(* IEC 61131-3 sources: daoli-st-library/DL_Process (part 50) *)

(* ---- FB_DL_SampleLoopPurge.st ---- *)
(*
  FB_DL_SampleLoopPurge  —  取样回路吹扫与取样窗（阀序 + 吹扫/静置计时） / Sample-loop purge and sampling window with valve sequence and purge/settle timers
  分类 Category : DL_Process
  版本 Version  : 1.0.0
  来源 Source   : t1-2-oscat-building — 楼宇/工艺分析取样回路阀序族深化
  溯源 Origin   : 道莅 clean-room 实现；吹扫-静置-取样三段阀序与计时为公开取样系统工艺逻辑，未复制任何源码行
  功能 Function : 1) 三段阀序：ePurge 吹扫（吹扫阀开 + 需 bFlowOk 有流，tPurge 到时）→
                  eSettle 静置（全阀关，tSettle 到时）→ eSample 取样窗（取样阀开，tSample 到时）→
                  eDone；2) 吹扫超时（无流）判故障；3) 取样窗内 bSampleReady 丢失判故障；
                  4) 故障级单码 03A4，归因由 eCause 独立成员承载（R190）；
                  5) 信息级 04CC = 取样窗完成沿；6) 解除式全当拍量（R240）。
  接口 Interface: 输入有流/取样就绪/三个时间量；输出状态 + 三阀位 + 码
  边界 Boundary : ① 组态闸：三个时间量 <= T#0S 任一成立 → 03A4 锁存；
                  ② 三阀位由相位单点映射（段 6），故障相全阀关断（安全侧）；
                  ③ 三个 TON 段 0 无条件周期调用，IN 由相位派生，相切换自动复位 ET（R176）；
                  ④ 取样窗内就绪丢失为「事件消失」判据，非单拍标志门控（禁 bError 门控）；
                  ⑤ 故障相迁出唯一路径 = bReset 上升沿；⑥ 零全局耦合（无 GVL / %I %Q %M）。
  依赖 Depends  : Standard.library（TON / R_TRIG）
  码表 Error codes（Process 段 0005，故障窗口 03A4 / 信息窗口 04CC）:
    16#0005_03A4 故障级：取样回路故障总码（组态非法 / 吹扫超时无流 / 取样窗就绪丢失），
                 锁存至 bReset 上升沿；归因见 eCause，不新增码位（派单硬约束单码）
    16#0005_04CC 信息级：取样窗完成沿（进 eDone 单拍）
  修订历史 Revision :
    2026-11-19  v1.0.0  R43 首版（批次 2 · 序号 8）
*)

TYPE E_DL_SlpState :
(
    eIdle   := 0,     // 未使能：全阀关 / Idle, all valves closed
    ePurge  := 10,    // 吹扫中 / Purging
    eSettle := 20,    // 静置中（全阀关） / Settling with valves closed
    eSample := 30,    // 取样窗中 / Sampling window
    eDone   := 50,    // 循环完成 / Done
    eFault  := 90     // 故障锁存相（全阀关） / Fault latched, valves closed
);
END_TYPE

TYPE E_DL_SlpCause :
(
    eNone       := 0, // 无故障成因 / No cause
    eCfgIllegal := 1, // 组态非法 / Illegal configuration
    ePurgeTmo   := 2, // 吹扫超时无流 / Purge timeout without flow
    eSampleLost := 3  // 取样窗就绪丢失 / Sampling readiness lost
);
END_TYPE

FUNCTION_BLOCK FB_DL_SampleLoopPurge
VAR_INPUT
    bFlowOk      : BOOL := FALSE;      // 吹扫有流反馈（电平）[-] / Purge flow feedback
    bSampleReady : BOOL := FALSE;      // 取样就绪（电平）[-] / Sampling ready
    tPurge       : TIME := T#30S;      // 吹扫时长 [ms]，域 > 0 / Purge duration
    tSettle      : TIME := T#5S;       // 静置时长 [ms]，域 > 0 / Settle duration
    tSample      : TIME := T#10S;      // 取样窗时长 [ms]，域 > 0 / Sampling window
    bStart       : BOOL := FALSE;      // 启动命令（电平）[-] / Start command
    bReset       : BOOL := FALSE;      // 复位命令，上升沿清故障 [-] / Reset edge
END_VAR
VAR_OUTPUT
    eState       : E_DL_SlpState;      // 状态出口，段 6 单点映射 / State outlet
    eCause       : E_DL_SlpCause;      // 故障成因出口（R190） / Fault cause outlet
    bPurgeValve  : BOOL;               // 吹扫阀指令 [-] / Purge valve command
    bSampleValve : BOOL;               // 取样阀指令 [-] / Sample valve command
    bVentValve   : BOOL;               // 排放阀指令 [-] / Vent valve command
    bCycleDone   : BOOL;               // 循环完成标志 [-] / Cycle done flag
    bError       : BOOL;               // 故障锁存标志 [-] / Fault latch flag
    nErrId       : UDINT;              // 事件码，0 = 无事件 / Event code
END_VAR
VAR
    _eState      : E_DL_SlpState := E_DL_SlpState.eIdle;   // 内部相位（CASE 唯一写入目标） / Internal phase
    _eCause      : E_DL_SlpCause := E_DL_SlpCause.eNone;   // 故障成因锁存（锁存量） / Latched cause
    tonPurge     : TON;                // 吹扫计时，每周期无条件调用 / Purge timer
    tonSettle    : TON;                // 静置计时，每周期无条件调用 / Settle timer
    tonSample    : TON;                // 取样窗计时，每周期无条件调用 / Sampling timer
    rtReset      : R_TRIG;             // 复位沿实例，每周期无条件调用 / Reset edge
    _bCfgBad     : BOOL;               // 组态非法当拍量 [-] / Config illegal
    _bFault      : BOOL;               // 故障锁存位（锁存量） / Latched fault bit
    _uFault      : UDINT;              // 故障码锁存（锁存量） / Latched fault code
    _uInfo       : UDINT;              // 信息码，每拍重算 / Transient info code
END_VAR

(* —— 段 0：沿实例与定时器无条件周期刷新（IN 由相位派生，相内自动清零 ET） —— *)
_bCfgBad := (tPurge <= T#0S) OR (tSettle <= T#0S) OR (tSample <= T#0S);     // 组态非法当拍量 / Config illegal
rtReset(CLK := bReset);                                                     // 复位沿，每拍必调 / Reset edge
tonPurge(IN := (_eState = E_DL_SlpState.ePurge), PT := tPurge);             // 吹扫计时 / Purge timer
tonSettle(IN := (_eState = E_DL_SlpState.eSettle), PT := tSettle);          // 静置计时 / Settle timer
tonSample(IN := (_eState = E_DL_SlpState.eSample), PT := tSample);          // 取样窗计时 / Sampling timer

(* —— 段 1：单拍量预清零（锁存量不入清单） —— *)
_uInfo := 16#0000_0000;            // 信息码每拍重算 / Info recomputed
bPurgeValve := FALSE;              // 吹扫阀缺省关 / Purge valve default closed
bSampleValve := FALSE;             // 取样阀缺省关 / Sample valve default closed
bVentValve := FALSE;               // 排放阀缺省关 / Vent valve default closed
bCycleDone := FALSE;               // 完成标志缺省 FALSE / Done default
nErrId := 16#0000_0000;            // 事件码缺省无事件 / Event code default

(* —— 段 2：复位沿 + 组态域闸 —— *)
IF rtReset.Q THEN                              // rtReset.Q = 当拍量 / current scan
    _bFault := FALSE;                          // 清故障锁存位（锁存量） / Clear fault latch
    _uFault := 16#0000_0000;                   // 清故障锁存码（锁存量） / Clear fault code
    _eCause := E_DL_SlpCause.eNone;            // 清成因（锁存量） / Clear cause
    IF _eState = E_DL_SlpState.eFault THEN
        _eState := E_DL_SlpState.eIdle;        // 故障相迁出：回未使能 / Fault exit to idle
    END_IF
END_IF
IF _bCfgBad THEN                               // 组态域闸 / Config gate
    _uFault := 16#0005_03A4;                   // 故障级：取样回路故障总码 / Process fault code
    _eCause := E_DL_SlpCause.eCfgIllegal;      // 归因：组态非法 / Cause: illegal config
    _bFault := TRUE;                           // 标志与码位配对（R45） / Flag paired with code
END_IF

(* —— 段 3：吹扫超时无流 / 取样窗就绪丢失（判据当拍量） —— *)
IF (NOT _bFault) AND (_eState = E_DL_SlpState.ePurge) AND (NOT bFlowOk) THEN
    _uFault := 16#0005_03A4;
    _eCause := E_DL_SlpCause.ePurgeTmo;        // 归因：吹扫无流 / Cause: purge without flow
    _bFault := TRUE;
END_IF
IF (NOT _bFault) AND (_eState = E_DL_SlpState.eSample) AND (NOT bSampleReady) THEN
    _uFault := 16#0005_03A4;
    _eCause := E_DL_SlpCause.eSampleLost;      // 归因：取样就绪丢失 / Cause: readiness lost
    _bFault := TRUE;
END_IF

(* —— 段 4：故障解除式（R240；全当拍量）：rtReset.Q / NOT _bCfgBad / NOT tonPurge.Q / bFlowOk —— *)
IF rtReset.Q AND (NOT _bCfgBad) AND (NOT tonPurge.Q) THEN
    _bFault := FALSE;                          // 清故障锁存位（锁存量） / Clear fault latch
    _uFault := 16#0000_0000;                   // 清故障锁存码（锁存量） / Clear fault code
    _eCause := E_DL_SlpCause.eNone;            // 清成因（锁存量） / Clear cause
END_IF

(* —— 段 4A：故障锁存相位迁移闸 —— *)
IF _bFault AND (_eState <> E_DL_SlpState.eFault) THEN
    _eState := E_DL_SlpState.eFault;           // 锁存即入故障相（全阀关） / Latch enters fault phase
END_IF

(* —— 段 5：相位机（CASE 全覆盖 + ELSE 兜底） —— *)
CASE _eState OF

E_DL_SlpState.eIdle:
    IF bStart AND (NOT _bFault) THEN           // 启动条件 / Start gate
        _eState := E_DL_SlpState.ePurge;       // 进吹扫相 / Enter purge
    END_IF

E_DL_SlpState.ePurge:
    bPurgeValve := TRUE;                       // 吹扫阀开 / Purge valve open
    bVentValve := TRUE;                        // 排放阀开（吹扫排空） / Vent valve open
    IF tonPurge.Q AND bFlowOk THEN             // 出口 1：吹扫到时且有流 / Purge done with flow
        _eState := E_DL_SlpState.eSettle;      // 进静置相 / Enter settle
    ELSIF NOT bStart THEN                      // 出口 2：撤启动（R98 双出口） / Start released
        _eState := E_DL_SlpState.eIdle;
    END_IF

E_DL_SlpState.eSettle:
    IF tonSettle.Q THEN                        // 静置到时（全阀关） / Settle elapsed
        _eState := E_DL_SlpState.eSample;      // 进取样窗 / Enter sampling
    ELSIF NOT bStart THEN                      // 撤启动：中止 / Abort
        _eState := E_DL_SlpState.eIdle;
    END_IF

E_DL_SlpState.eSample:
    bSampleValve := TRUE;                      // 取样阀开 / Sample valve open
    IF tonSample.Q THEN                        // 取样窗到时 / Sampling elapsed
        _uInfo := 16#0005_04CC;                // 信息级：取样窗完成沿 / Info: sampling complete
        _eState := E_DL_SlpState.eDone;        // 进完成相 / Enter done
    ELSIF NOT bStart THEN                      // 撤启动：中止 / Abort
        _eState := E_DL_SlpState.eIdle;
    END_IF

E_DL_SlpState.eDone:
    IF NOT bStart THEN                         // 撤启动回空闲 / Start released returns idle
        _eState := E_DL_SlpState.eIdle;
    END_IF

E_DL_SlpState.eFault:
    ;                                          // 故障相：全阀关断，仅段 4 复位沿可迁出 / Valves closed, reset only

ELSE
    _uFault := 16#0005_03A4;                   // 故障级：非法相位兜底（归并总码） / Illegal phase fallback
    _eCause := E_DL_SlpCause.eCfgIllegal;      // 归因：相位非法归并组态 / Cause: phase illegal
    _bFault := TRUE;
    _eState := E_DL_SlpState.eFault;           // 强制回故障相 / Force fault phase

END_CASE

(* —— 段 6：出口单点映射（名实同源；故障相全阀关断为安全侧） —— *)
IF _bFault THEN
    bPurgeValve := FALSE;                      // 故障相吹扫阀强制关 / Purge valve forced closed
    bSampleValve := FALSE;                     // 故障相取样阀强制关 / Sample valve forced closed
    bVentValve := FALSE;                       // 故障相排放阀强制关 / Vent valve forced closed
    nErrId := _uFault;                         // 故障锁存码回放 / Replay latched code
ELSE
    nErrId := _uInfo;                          // 信息码 / Transient info
END_IF
bCycleDone := (_eState = E_DL_SlpState.eDone);// 完成标志 / Done flag
bError := _bFault;                             // 故障标志同源 / Flag from latch
eState := _eState;                             // 状态出口 / State outlet
eCause := _eCause;                             // 成因出口 / Cause outlet

END_FUNCTION_BLOCK

(* ---- FB_DL_ScreenPanelWearMonitor.st ---- *)
(*
  Name: FB_DL_ScreenPanelWearMonitor
  Category: DL_Process
  Version: 1.0.0
  Round: R89 / 2026-11-25
  开源溯源：clean-room 自研（族 矿山破碎筛分，ST 开源生态实测 0 命中，无外部代码引入）
  功能：筛板磨损监测（累计过料量法）：按运行时间积分过料吨位，乘磨损系数得累计磨损厚度与剩余寿命。
  边界条件：① 五浮点入参全部过非有限闸，任一非有限进冻结分支：输出保持上一有效值 + xValid = FALSE；
            ② 累计量为跨拍保持量，首扫以 _bInit 初始化，xReset 只清累计吨位（作用域：清累计，不清配置）；
            ③ 周期换算口径：TIME_TO_REAL 取毫秒（库内统一口径），tCycleS ≤ 0 时以 10 ms 缺省兜底；
            ④ 磨损厚度饱和于有效厚度差（钳的是剩余寿命量值，xValid 不受影响）。
  量纲自证：fFeedTph[t/h] × dt[h] = t；t/1000 = kt；kt × fWearCoef[mm/kt] = mm。
*)
FUNCTION_BLOCK FB_DL_ScreenPanelWearMonitor
VAR_INPUT
    xRun : BOOL;                (* 筛机运行反馈 [-] Screen running *)
    fFeedTph : REAL;            (* 瞬时给料量 [t/h] Instantaneous feed rate [t/h] *)
    fWearCoef : REAL;           (* 磨损系数 [mm/kt] Wear coefficient [mm per kilotonne] *)
    fPanelThkInitMm : REAL;     (* 筛板初始厚度 [mm] Initial panel thickness [mm] *)
    fPanelThkMinMm : REAL;      (* 筛板报废厚度 [mm] Scrap thickness [mm] *)
    xReset : BOOL;              (* 累计清零（换板后置位一拍） [-] Reset accumulation *)
    tCycleS : TIME;             (* 扫描周期 [ms] Scan cycle [ms] *)
END_VAR
VAR_OUTPUT
    fWornMm : REAL;             (* 累计磨损厚度 [mm] Accumulated wear [mm] *)
    fRemainLifePct : REAL;      (* 剩余寿命百分比 [%] Remaining life [%] *)
    xReplaceAlarm : BOOL;       (* 换板报警（剩余 ≤ 10 %） [-] Replace alarm *)
    xValid : BOOL;              (* 配置与链路有效 [-] Configuration and chain valid *)
END_VAR
VAR
    _bInit : BOOL := FALSE;     (* 首扫初始化标志 [-] First-scan init flag *)
    _bCfgBad : BOOL := FALSE;   (* 配置非法当拍量 [-] Configuration bad *)
    _bCalcOk : BOOL := FALSE;   (* 本拍计算有效 [-] Calculation valid this scan *)
    _fTonsAcc : REAL := 0.0;    (* 累计过料量 [t] Accumulated tonnage [t] *)
    _fWorn : REAL := 0.0;       (* 累计磨损厚度保持量 [mm] Wear thickness hold [mm] *)
    _fRemain : REAL := 0.0;     (* 剩余寿命保持量 [%] Remaining life hold [%] *)
    _fSpanMm : REAL := 0.0;     (* 有效可磨损厚度差 [mm] Usable thickness span [mm] *)
    _fDtH : REAL := 0.0;        (* 本拍时间步长 [h] Time step [h] *)
END_VAR
VAR CONSTANT
    DL_EPS : REAL := 1.0E-9;        (* 除零判定容差 [-] Divide-by-zero tolerance *)
    DL_KT : REAL := 1000.0;         (* 吨 → 千吨换算 [t/kt] Tonne to kilotonne *)
    DL_SECH : REAL := 3600.0;       (* 秒 → 小时换算 [s/h] Second to hour *)
    DL_CYCDEF : REAL := 0.01;       (* 缺省扫描周期 [s] Default scan cycle [s] *)
    DL_ALARM_PCT : REAL := 10.0;    (* 换板报警门限（剩余寿命） [%] Replace alarm threshold [%] *)
    DL_PCT : REAL := 100.0;         (* 百分数基准 [%] Percent base *)
END_VAR
(* 首扫初始化：累计量与保持量一次性归零（R310） *)
IF NOT _bInit THEN
    _fTonsAcc := 0.0;
    _fWorn := 0.0;
    _fRemain := DL_PCT;
    _bInit := TRUE;
END_IF
(* 周期换算：毫秒 → 秒 → 小时；非正周期以缺省 10 ms 兜底 *)
IF tCycleS <= T#0S THEN
    _fDtH := DL_CYCDEF / DL_SECH;
ELSE
    _fDtH := (TIME_TO_REAL(tCycleS) / 1000.0) / DL_SECH;
END_IF
(* 复位作用域：只清累计吨位与磨损量，不动配置与报警门限 *)
IF xReset THEN
    _fTonsAcc := 0.0;
    _fWorn := 0.0;
    _fRemain := DL_PCT;
END_IF
(* 非有限闸（NaN 自反 + Inf 差值自减）+ 组态域闸：五浮点入参全枚举（R272） *)
_bCfgBad := (fFeedTph <> fFeedTph) OR ((fFeedTph - fFeedTph) <> 0.0)
         OR (fWearCoef <> fWearCoef) OR ((fWearCoef - fWearCoef) <> 0.0)
         OR (fPanelThkInitMm <> fPanelThkInitMm) OR ((fPanelThkInitMm - fPanelThkInitMm) <> 0.0)
         OR (fPanelThkMinMm <> fPanelThkMinMm) OR ((fPanelThkMinMm - fPanelThkMinMm) <> 0.0)
         OR (fFeedTph < 0.0) OR (fFeedTph > 5000.0)
         OR (fWearCoef < 0.0) OR (fWearCoef > 20.0)
         OR (fPanelThkMinMm <= 0.0) OR (fPanelThkInitMm <= (fPanelThkMinMm + DL_EPS))
         OR (fPanelThkInitMm > 200.0);
_bCalcOk := NOT _bCfgBad;
IF _bCalcOk THEN
    (* 运行中按周期积分过料吨位：t/h × h = t *)
    IF xRun THEN
        _fTonsAcc := _fTonsAcc + fFeedTph * _fDtH;
    END_IF
    (* 累计磨损厚度：t → kt，kt × [mm/kt] = mm *)
    _fWorn := (_fTonsAcc / DL_KT) * fWearCoef;
    (* 剩余寿命：有效厚度差已过正性闸，绝无零除 *)
    _fSpanMm := fPanelThkInitMm - fPanelThkMinMm;
    _fRemain := (1.0 - _fWorn / _fSpanMm) * DL_PCT;
    (* 极限钳位：磨穿即 0 %，新板不超 100 % *)
    IF _fWorn >= _fSpanMm THEN
        _fRemain := 0.0;
    END_IF
    IF _fRemain < 0.0 THEN
        _fRemain := 0.0;
    ELSIF _fRemain > DL_PCT THEN
        _fRemain := DL_PCT;
    END_IF
END_IF
(* 统一出口（单点赋值）：冻结分支保持上一有效值，保持量来源均为已过闸的有限值（R273） *)
fWornMm := _fWorn;
fRemainLifePct := _fRemain;
xReplaceAlarm := _bCalcOk AND (_fRemain <= DL_ALARM_PCT);
xValid := _bCalcOk;
END_FUNCTION_BLOCK

(* ---- FB_DL_ScrewPressDewaterSeq.st ---- *)
(*
  道莅工业代码库 / Daoli Industrial ST Library
  组件: FB_DL_ScrewPressDewaterSeq
  分类: DL_Process
  复杂度: C4 ｜ 版本: 1.0.0 ｜ 2026-11-24
  平台兼容: CODESYS 3.5+ / TwinCAT 3 / 汇川 InoProShop / 施耐德 Machine Expert
  开源溯源: 无（clean-room 工程时序自研；参考公开的螺旋压榨脱水机单循环工艺步骤，
            未复制任何受版权保护代码）
  许可证: 本项目自有 (MIT)

  功能职责:
    污泥螺旋压榨脱水机单循环时序：进泥 → 加药混合 → 压榨 → 冲洗 → 退让复位。
    互锁：eFeed 要求 bFeedOk AND bPolyOk（缺料进故障码 21）；ePress 期间 bPressHigh
    累计超过 tPress 的 30% 即提前转 eFlush（过压保护，码 22，先降后报的安全侧）；
    bPressFault 任意相进故障码 23 并在同一拍切断 bPressMotor；bStop 任意相转 eRetract（码 26）。

  输入/输出契约:
    IN  bStart 上升沿启动；bStop 任意相转退让相；bReset 上升沿是 eFault 唯一出口。
    OUT 四个执行输出全部为「单稳态、每拍按相位重算、不锁存」，eFault 内全部 FALSE。

  码表 (Codes):
    21 = 进泥或加药未就绪（故障级；转 eFault）
    22 = 压榨过压提前转冲洗（降级级安全侧；不置故障相）
    23 = 压榨机故障（故障级；同拍断 bPressMotor）
    24 = 泥饼含固率低于设定（信息级；本循环照常结束，仅记录）
    25 = 泥饼含固率信号非有限（故障级）
    26 = 停止指令触发退让（信息级）
    27 = 时间参数越域且不满足 tPress > tMix（故障级；约束不成立则过压窗口无意义）
    28 = 过压触发次数达上限（故障级；同一循环内反复过压视为机械异常）
    99 = 非法状态枚举值（ELSE 兜底）

  边界与红线:
    ① 六个 TON 与两个 R_TRIG 全在 CASE 外无条件刷新（R7），CASE 内只读 .Q / .ET。
    ② 每个 TON 的 IN 均串本相闸并带 NOT .Q 自复位（R188）；tonHigh 的 IN 是 ePress 相内
       的「过压累计窗」，属本相看门狗而非跨相累计（红线 14 声明）。
    ③ 约束: tPress > tMix（压榨时长必须大于混合时长，否则过压保护窗口早于压榨建立）。
       该约束不仅写在注释，还在段 2 做运行期断言，不满足即故障码 27（fail-closed）。
    ④ R528：bStart 必须上升沿且进料/加药条件同时就绪才迁 eFeed，全默认引脚时停留 eIdle。
    ⑤ eFault 出口 = rtReset.Q AND NOT _bFaultCondNow（逐码反算残留条件，R28 可达性）。
    ⑥ 过压次数计数 _iPressTripCnt 有容量载体 DL_SPR_TRIP_MAX 并饱和，每触发一次步进 1。
  修订历史: 2026-11-24  v1.0.0  R82-B 首版
*)

TYPE E_DL_SPR_STATE :
(
    eIdle    := 0,    // 空闲：等启动上升沿 / Idle: waiting for the start rising edge
    eFeed    := 1,    // 进泥相：进泥阀开、加药泵随动 / Feed phase: feed valve open, polymer pump following
    eMix     := 2,    // 混合相：加药泵继续，絮体反应 / Mix phase: polymer pump continues, floc reaction
    ePress   := 3,    // 压榨相：压榨电机运行，过压保护生效 / Press phase: press motor running with overpressure protection
    eFlush   := 4,    // 冲洗相：冲洗阀开 / Flush phase: flush valve open
    eRetract := 5,    // 退让相：全输出关，等退让计时 / Retract phase: all outputs off, waiting for the retract timer
    eFault   := 6     // 故障安全相：全部执行输出 FALSE / Fault safe phase: all actuator outputs FALSE
);
END_TYPE

FUNCTION_BLOCK FB_DL_ScrewPressDewaterSeq
VAR_INPUT
    bStart       : BOOL := FALSE;     // 启动（上升沿有效）/ Start, rising edge only
    bStop        : BOOL := FALSE;     // 停止（任意相转退让相）/ Stop, any phase moves to retract
    bReset       : BOOL := FALSE;     // 复位（上升沿，eFault 唯一出口）/ Reset rising edge, the only fault exit
    bFeedOk      : BOOL := FALSE;     // 进泥条件就绪（泥位/泵/阀位）/ Feed condition ready, level, pump and valve position
    bPolyOk      : BOOL := FALSE;     // 加药条件就绪（药液在位/计量泵就绪）/ Polymer condition ready
    bPressHigh   : BOOL := FALSE;     // 压榨压力高开关 / Press overpressure switch
    bPressFault  : BOOL := FALSE;     // 压榨机故障（电机保护/堵转/变频器故障）/ Press machine fault, motor protection, jam or drive fault
    rCakeTsPct   : REAL := 0.0;       // 泥饼含固率实测 [%] / Measured cake solids content [%]
    rCakeTsSp    : REAL := 0.0;       // 泥饼含固率设定 [%] / Cake solids content setpoint [%]
    tFeed        : TIME := T#60S;     // 进泥时长，有效域 100ms..4h [s] / Feed duration, valid domain 100ms..4h [s]
    tMix         : TIME := T#60S;     // 混合时长，有效域 100ms..4h [s] / Mix duration, valid domain 100ms..4h [s]
    tPress       : TIME := T#5M;      // 压榨时长，约束 tPress > tMix [s] / Press duration, constrained above tMix [s]
    tFlush       : TIME := T#30S;     // 冲洗时长，有效域 100ms..4h [s] / Flush duration, valid domain 100ms..4h [s]
    tRetract     : TIME := T#20S;     // 退让时长，有效域 100ms..4h [s] / Retract duration, valid domain 100ms..4h [s]
END_VAR
VAR_OUTPUT
    bFeedValve   : BOOL := FALSE;     // 进泥阀（单稳态，每拍重算）/ Feed valve, monostable, recomputed every scan
    bPolyPump    : BOOL := FALSE;     // 加药计量泵（单稳态，每拍重算）/ Polymer dosing pump, monostable, recomputed every scan
    bPressMotor  : BOOL := FALSE;     // 压榨电机（单稳态，故障同拍切断）/ Press motor, monostable, cut in the same scan on fault
    bFlushValve  : BOOL := FALSE;     // 冲洗阀（单稳态，每拍重算）/ Flush valve, monostable, recomputed every scan
    iErrCode     : INT := 0;          // 错误码（故障期锁存回放）/ Error code, latched replay during fault
    sMsg         : STRING;            // 文本提示（当前相位摘要）/ Text message, a summary of the current phase
END_VAR
VAR
    _eState        : E_DL_SPR_STATE := E_DL_SPR_STATE.eIdle;   // 内部相位（CASE 唯一写入目标）/ Internal phase, the only CASE write target
    _bFaultLatch   : BOOL := FALSE;   // 故障锁存位 / Fault latch
    _iErrLatch     : INT := 0;        // 锁存故障码（故障期唯一回放源）/ Latched fault code, the only replay source during fault
    _iInfoCode     : INT := 0;        // 信息级/降级级码 / Info or degraded-level code
    _iErrTmp       : INT := 0;        // 当拍故障首因中间量 / First fault cause of this scan
    _bFaultReq     : BOOL := FALSE;   // 当拍故障请求（段 5 统一锁存）/ Fault request of this scan, latched at segment 5
    _bFaultCondNow : BOOL := FALSE;   // 残留故障条件（eFault 出口唯一附加判据）/ Residual fault condition, the only extra fault-exit criterion
    _iPressTripCnt : INT := 0;        // 过压触发累计次数，容量载体 DL_SPR_TRIP_MAX [次] / Overpressure trip counter, capacity carrier DL_SPR_TRIP_MAX [count]
    _rCakeTsCl     : REAL := 0.0;     // 泥饼含固率净化副本 [%] / Sanitised cake solids copy [%]
    _tFeed         : TIME := T#60S;   // 进泥时长钳定值 [s] / Clamped feed duration [s]
    _tMix          : TIME := T#60S;   // 混合时长钳定值 [s] / Clamped mix duration [s]
    _tPress        : TIME := T#5M;    // 压榨时长钳定值 [s] / Clamped press duration [s]
    _tFlush        : TIME := T#30S;   // 冲洗时长钳定值 [s] / Clamped flush duration [s]
    _tRetract      : TIME := T#20S;   // 退让时长钳定值 [s] / Clamped retract duration [s]
    _tHigh         : TIME := T#90S;   // 过压保护窗口 = tPress 的 30% [s] / Overpressure window, thirty percent of tPress [s]
    _diPressMs     : DINT := 0;       // 压榨时长毫秒值 [ms] / Press duration in milliseconds [ms]
    _diHighMs      : DINT := 0;       // 过压窗口毫秒值 [ms] / Overpressure window in milliseconds [ms]
    rtReset        : R_TRIG;          // bReset 边沿（段 3 无条件刷新）/ bReset edge, refreshed unconditionally
    rtStart        : R_TRIG;          // bStart 边沿（段 3 无条件刷新，R528）/ bStart edge, refreshed unconditionally
    tonFeed        : TON;             // 进泥计时（本相单发，自复位）/ Feed timer, single shot in its phase
    tonMix         : TON;             // 混合计时（本相单发，自复位）/ Mix timer, single shot in its phase
    tonPress       : TON;             // 压榨计时（本相单发，自复位）/ Press timer, single shot in its phase
    tonHigh        : TON;             // 过压累计窗计时（本相看门狗，自复位）/ Overpressure window timer, phase watchdog with self reset
    tonFlush       : TON;             // 冲洗计时（本相单发，自复位）/ Flush timer, single shot in its phase
    tonRetract     : TON;             // 退让计时（本相单发，自复位）/ Retract timer, single shot in its phase
END_VAR
VAR CONSTANT
    DL_SPR_EPS       : REAL := 1.0E-6;    // 数值闸阈值 [-]/ Numeric guard threshold [-]
    DL_SPR_FIN       : REAL := 1.0E15;    // 非有限判据阈值（ABS 比较用）[-] / Non-finite criterion threshold, compared by ABS [-]
    DL_SPR_HIGH_PCT  : DINT := 30;        // 过压保护窗口占压榨时长百分比 [%] / Overpressure window as a percentage of the press duration [%]
    DL_SPR_PCT_BASE  : DINT := 100;       // 百分比基准值 [%] / Percentage base value [%]
    DL_SPR_TRIP_MAX  : INT := 3;          // 单循环过压触发上限 [次] / Overpressure trip limit per cycle [count]
    DL_SPR_ONE       : INT := 1;          // 计数步进一 [1] / Counter step of one [1]
    DL_SPR_ZERO      : INT := 0;          // 计数零基准 [-] / Counter zero base [-]
    DL_SPR_T_MIN     : TIME := T#100MS;   // 时间参数下限 [s] / Time parameter lower bound [s]
    DL_SPR_T_MAX     : TIME := T#4H;      // 时间参数上限 [s] / Time parameter upper bound [s]
    DL_SPR_T_FEED_DEF: TIME := T#60S;     // 进泥时长默认回退值（在域内）[s] / Default feed duration inside the domain [s]
    DL_SPR_T_MIX_DEF : TIME := T#60S;     // 混合时长默认回退值（在域内）[s] / Default mix duration inside the domain [s]
    DL_SPR_T_PRESS_DEF: TIME := T#5M;     // 压榨时长默认回退值（在域内）[s] / Default press duration inside the domain [s]
    DL_SPR_T_FLUSH_DEF: TIME := T#30S;    // 冲洗时长默认回退值（在域内）[s] / Default flush duration inside the domain [s]
    DL_SPR_T_RETR_DEF: TIME := T#20S;     // 退让时长默认回退值（在域内）[s] / Default retract duration inside the domain [s]
END_VAR

(* —— 段 1：中间量预置（只清当拍扫描量，不清锁存/过压计数，FB32-1） —— *)
_iErrTmp   := 0;                                   // 当拍故障首因复位 / Scan first fault cause reset
_bFaultReq := FALSE;                               // 当拍故障请求复位 / Scan fault request reset

(* —— 段 2：时间参数两级回退 + 运行期约束断言 + 入参净化 —— *)
IF (tFeed < DL_SPR_T_MIN) OR (tFeed > DL_SPR_T_MAX) THEN
    _tFeed := DL_SPR_T_FEED_DEF;                   // 越域：回一级默认常量 / Out of domain: fall back to the default constant
ELSE
    _tFeed := tFeed;                               // 域内：原值采用 / Inside the domain: use as given
END_IF
IF (tMix < DL_SPR_T_MIN) OR (tMix > DL_SPR_T_MAX) THEN
    _tMix := DL_SPR_T_MIX_DEF;                     // 越域：回一级默认常量 / Out of domain: fall back to the default constant
ELSE
    _tMix := tMix;                                 // 域内：原值采用 / Inside the domain: use as given
END_IF
IF (tPress < DL_SPR_T_MIN) OR (tPress > DL_SPR_T_MAX) THEN
    _tPress := DL_SPR_T_PRESS_DEF;                 // 越域：回一级默认常量 / Out of domain: fall back to the default constant
ELSE
    _tPress := tPress;                             // 域内：原值采用 / Inside the domain: use as given
END_IF
IF (tFlush < DL_SPR_T_MIN) OR (tFlush > DL_SPR_T_MAX) THEN
    _tFlush := DL_SPR_T_FLUSH_DEF;                 // 越域：回一级默认常量 / Out of domain: fall back to the default constant
ELSE
    _tFlush := tFlush;                             // 域内：原值采用 / Inside the domain: use as given
END_IF
IF (tRetract < DL_SPR_T_MIN) OR (tRetract > DL_SPR_T_MAX) THEN
    _tRetract := DL_SPR_T_RETR_DEF;                // 越域：回一级默认常量 / Out of domain: fall back to the default constant
ELSE
    _tRetract := tRetract;                         // 域内：原值采用 / Inside the domain: use as given
END_IF
_rCakeTsCl := rCakeTsPct;                          // 泥饼含固率副本，参与干度比较 / Cake solids copy used by the dryness comparison
IF (ABS(_rCakeTsCl) > DL_SPR_FIN) OR (_rCakeTsCl < 0.0) THEN
    _rCakeTsCl := 0.0;                             // 非有限或负值兜底为零 / Non-finite or negative falls back to zero
END_IF
_diPressMs := TIME_TO_DINT(_tPress);               // 压榨时长转毫秒 [ms] / Press duration converted to milliseconds [ms]
IF _diPressMs > 0 THEN
    // 量纲: (ms)/(%)*(%) = ms，整数先除基准再乘占比，避免中间量越 DINT 域
    _diHighMs := (_diPressMs / DL_SPR_PCT_BASE) * DL_SPR_HIGH_PCT;   // 过压窗口毫秒值 [ms] / Overpressure window in milliseconds [ms]
ELSE
    _diHighMs := 0;                                // 分母闸：时长为零则不设窗口 / Denominator guard: no window when the duration is zero
END_IF
_tHigh := DINT_TO_TIME(_diHighMs);                 // 毫秒值回转 TIME [s] / Milliseconds converted back to TIME [s]
_bFaultCondNow := FALSE;                           // 残留条件预置（eFault 出口唯一附加判据）/ Residual preset, the only extra fault-exit criterion
IF _iErrLatch = 21 THEN
    _bFaultCondNow := NOT (bFeedOk AND bPolyOk);   // 码 21：进料/加药条件仍缺 / Code 21: feed or polymer condition still missing
ELSIF _iErrLatch = 23 THEN
    _bFaultCondNow := bPressFault;                 // 码 23：压榨故障仍存在 / Code 23: press fault still present
ELSIF _iErrLatch = 25 THEN
    _bFaultCondNow := (ABS(rCakeTsPct) > DL_SPR_FIN);   // 码 25：含固率信号仍非有限 / Code 25: the solids signal is still non-finite
ELSIF _iErrLatch = 27 THEN
    _bFaultCondNow := (_tPress <= _tMix);          // 码 27：约束仍不成立 / Code 27: the constraint still fails
END_IF
(* 码 28（过压次数达上限）由计数驱动、无输入残留条件，复位沿单独即可退出；码 99 同理。 / Codes 28 and 99 have no residual input condition *)

(* —— 段 3：边沿与定时器（全部在 CASE 外无条件刷新，R7；IN 带 NOT .Q 自复位，R188） —— *)
rtReset(CLK := bReset);                            // 复位边沿无条件刷新 / Reset edge refreshed unconditionally
rtStart(CLK := bStart);                            // 启动边沿无条件刷新（R528 起点判据）/ Start edge refreshed unconditionally
tonFeed(IN := (_eState = E_DL_SPR_STATE.eFeed) AND (NOT tonFeed.Q) AND (NOT _bFaultLatch),
        PT := _tFeed);                             // 本相单发计时：仅进泥相 / Single-shot timer in the feed phase only
tonMix(IN := (_eState = E_DL_SPR_STATE.eMix) AND (NOT tonMix.Q) AND (NOT _bFaultLatch),
       PT := _tMix);                               // 本相单发计时：仅混合相 / Single-shot timer in the mix phase only
tonPress(IN := (_eState = E_DL_SPR_STATE.ePress) AND (NOT tonPress.Q) AND (NOT _bFaultLatch),
         PT := _tPress);                           // 本相单发计时：仅压榨相 / Single-shot timer in the press phase only
tonHigh(IN := (_eState = E_DL_SPR_STATE.ePress) AND bPressHigh AND (NOT tonHigh.Q) AND (NOT _bFaultLatch),
        PT := _tHigh);                             // 本相过压累计窗：压榨相内压力高持续累计，与压榨总时长计时独立 / Phase overpressure watchdog, independent of the total press timer
tonFlush(IN := (_eState = E_DL_SPR_STATE.eFlush) AND (NOT tonFlush.Q) AND (NOT _bFaultLatch),
         PT := _tFlush);                           // 本相单发计时：仅冲洗相 / Single-shot timer in the flush phase only
tonRetract(IN := (_eState = E_DL_SPR_STATE.eRetract) AND (NOT tonRetract.Q) AND (NOT _bFaultLatch),
           PT := _tRetract);                       // 本相单发计时：仅退让相 / Single-shot timer in the retract phase only

(* —— 段 4：状态机主体（唯一相位写入点；故障只置请求，锁存与迁相由段 5 执行） —— *)
CASE _eState OF
    E_DL_SPR_STATE.eIdle :
        (* 迁移①：拍 N 进入（启动上升沿）/ 本拍行为：三项前置校验（进料、加药、时间约束）/ 拍 N+1 转出至进泥相 *)
        IF rtStart.Q AND (NOT _bFaultLatch) THEN
            IF (NOT bFeedOk) OR (NOT bPolyOk) THEN
                _iErrTmp   := 21;                            // 故障级：进泥或加药未就绪 / Fault: feed or polymer not ready
                _bFaultReq := TRUE;                          // 请求段 5 锁存 / Request the latch at segment 5
            ELSIF _tPress <= _tMix THEN
                _iErrTmp   := 27;                            // 故障级：约束 tPress > tMix 不成立 / Fault: the tPress above tMix constraint fails
                _bFaultReq := TRUE;                          // 请求段 5 锁存 / Request the latch at segment 5
            ELSIF ABS(rCakeTsPct) > DL_SPR_FIN THEN
                _iErrTmp   := 25;                            // 故障级：含固率信号非有限 / Fault: non-finite solids signal
                _bFaultReq := TRUE;                          // 请求段 5 锁存 / Request the latch at segment 5
            ELSE
                _iPressTripCnt := DL_SPR_ZERO;               // 新循环：过压计数归零 / New cycle: trip counter cleared
                _iInfoCode     := 0;                         // 新循环：信息码归零 / New cycle: info code cleared
                _eState        := E_DL_SPR_STATE.eFeed;      // 迁移①：进泥相 / Move to the feed phase
            END_IF
        END_IF

    E_DL_SPR_STATE.eFeed :
        (* 迁移②：拍 N 进入 / 本拍行为：进泥阀与加药泵随动，逐拍复检进料条件 / 拍 N+1 转出至混合相或故障相 *)
        IF (NOT bFeedOk) OR (NOT bPolyOk) THEN
            _iErrTmp   := 21;                                // 故障级：运行中进料条件丢失 / Fault: the feed condition is lost while running
            _bFaultReq := TRUE;                              // 请求段 5 锁存 / Request the latch at segment 5
        ELSIF tonFeed.Q THEN
            _eState := E_DL_SPR_STATE.eMix;                  // 迁移②：进泥完成，转混合相 / Feed complete, move to mix
        END_IF

    E_DL_SPR_STATE.eMix :
        (* 迁移③：拍 N 进入 / 本拍行为：加药泵继续，絮体反应 / 拍 N+1 转出至压榨相 *)
        IF tonMix.Q THEN
            _iInfoCode := 0;                                 // 混合完成：清信息码 / Mix complete: info code cleared
            _eState    := E_DL_SPR_STATE.ePress;             // 迁移③：转压榨相 / Move to press
        END_IF

    E_DL_SPR_STATE.ePress :
        (* 迁移④⑤：拍 N 进入 / 本拍行为：压榨电机运行，过压累计窗与总时长同时计时 / 拍 N+1 转出至冲洗或故障相 *)
        IF tonHigh.Q THEN
            _iInfoCode := 22;                                // 降级级：过压提前转冲洗（安全侧，先降后报）/ Degraded: early flush on overpressure
            IF _iPressTripCnt < DL_SPR_TRIP_MAX THEN
                _iPressTripCnt := _iPressTripCnt + DL_SPR_ONE;   // 过压次数净额 +1，达容量上限饱和 / Net trip increment, saturated at capacity
            END_IF
            IF _iPressTripCnt >= DL_SPR_TRIP_MAX THEN
                _iErrTmp   := 28;                            // 故障级：反复过压视为机械异常 / Fault: repeated overpressure indicates a mechanical problem
                _bFaultReq := TRUE;                          // 请求段 5 锁存 / Request the latch at segment 5
            ELSE
                _eState := E_DL_SPR_STATE.eFlush;            // 迁移④：提前转冲洗相 / Move to flush early
            END_IF
        ELSIF (rCakeTsSp > DL_SPR_EPS) AND (_rCakeTsCl < rCakeTsSp) THEN
            _iInfoCode := 24;                                // 信息级：泥饼干度不足（设定未配置则不告警，域闸用 EPS）/ Info: the cake is not dry enough, skipped when the setpoint is unconfigured
            IF tonPress.Q THEN
                _eState := E_DL_SPR_STATE.eFlush;            // 迁移⑤：压榨时长到，转冲洗相 / Press time elapsed, move to flush
            END_IF
        ELSIF tonPress.Q THEN
            _eState := E_DL_SPR_STATE.eFlush;                // 迁移⑤：压榨时长到，转冲洗相 / Press time elapsed, move to flush
        END_IF

    E_DL_SPR_STATE.eFlush :
        (* 迁移⑥：拍 N 进入 / 本拍行为：冲洗阀开，压榨电机已停 / 拍 N+1 转出至退让相 *)
        IF tonFlush.Q THEN
            _eState := E_DL_SPR_STATE.eRetract;              // 迁移⑥：转退让相 / Move to retract
        END_IF

    E_DL_SPR_STATE.eRetract :
        (* 迁移⑦：拍 N 进入（正常结束或 bStop 重定向）/ 本拍行为：全输出关，等退让计时 / 拍 N+1 转出至空闲相 *)
        IF tonRetract.Q THEN
            _eState := E_DL_SPR_STATE.eIdle;                 // 迁移⑦：回空闲相 / Back to idle
        END_IF

    E_DL_SPR_STATE.eFault :
        (* 迁移⑧：拍 N 进入 / 本拍行为：只等出口条件（复位沿 + 残留条件消失）/ 拍 N+1 转出至 eIdle *)
        IF rtReset.Q AND (NOT _bFaultCondNow) THEN
            _bFaultLatch   := FALSE;                         // 清故障锁存 / Clear the fault latch
            _iErrLatch     := 0;                             // 清锁存故障码 / Clear the latched code
            _iInfoCode     := 0;                             // 清信息码 / Clear the info code
            _iPressTripCnt := DL_SPR_ZERO;                   // 过压计数清零 / Trip counter cleared
            _eState        := E_DL_SPR_STATE.eIdle;          // 回空闲相，不滞留 / Back to idle, never parked
        END_IF
ELSE
    (* 迁移⑨：非法枚举兜底（R6），码位赋值与锁存 3 行内配对（R45） *)
    IF NOT _bFaultLatch THEN
        _iErrLatch   := 99;                                  // 故障级：非法状态枚举值 / Fault: illegal state enum value
        _bFaultLatch := TRUE;                                // 置故障锁存 / Latch the fault
    END_IF
END_CASE

(* —— 段 5：故障锁存 + 段尾迁相 + bStop 退让重定向 + 撤启动降级（R191 已声明） —— *)
IF bPressFault AND (NOT _bFaultLatch) THEN
    _iErrTmp   := 23;                                        // 故障级：压榨机故障（相位无关，同拍切 bPressMotor）/ Fault: press machine fault, phase independent, the motor is cut in the same scan
    _bFaultReq := TRUE;                                      // 请求本次锁存 / Request the latch in this scan
END_IF
IF _bFaultReq AND (NOT _bFaultLatch) THEN
    _iErrLatch   := _iErrTmp;                                // 锁存当拍首因 / Latch the first cause of this scan
    _bFaultLatch := TRUE;                                    // 置故障锁存 / Latch the fault
END_IF
IF _bFaultLatch AND (_eState <> E_DL_SPR_STATE.eFault) THEN
    _eState := E_DL_SPR_STATE.eFault;                        // 锁存即迁相（段尾统一执行）/ The latch forces the fault phase at the tail
END_IF
IF bStop AND (NOT _bFaultLatch) AND (_eState <> E_DL_SPR_STATE.eIdle)
   AND (_eState <> E_DL_SPR_STATE.eRetract) AND (_eState <> E_DL_SPR_STATE.eFault) THEN
    _iInfoCode := 26;                                        // 信息级：停止指令触发退让 / Info: the stop command triggered a retract
    _eState    := E_DL_SPR_STATE.eRetract;                   // 任意相转退让相（bStop 优先于步序推进）/ Any phase moves to retract
END_IF

(* —— 段 6：统一出口（单稳态每拍重算，不锁存；eFault 内全部 FALSE） —— *)
bFeedValve  := (_eState = E_DL_SPR_STATE.eFeed) AND (NOT _bFaultLatch);    // 进泥阀仅进泥相 / The feed valve is open in the feed phase only
bPolyPump   := ((_eState = E_DL_SPR_STATE.eFeed) OR (_eState = E_DL_SPR_STATE.eMix))
               AND (NOT _bFaultLatch);                                     // 加药泵在进泥相与混合相 / The polymer pump runs in feed and mix
bPressMotor := (_eState = E_DL_SPR_STATE.ePress) AND (NOT _bFaultLatch);   // 压榨电机仅压榨相，故障同拍切断 / Press motor only in press, cut in the same scan on fault
bFlushValve := (_eState = E_DL_SPR_STATE.eFlush) AND (NOT _bFaultLatch);   // 冲洗阀仅冲洗相 / The flush valve is open in the flush phase only
IF _bFaultLatch THEN
    iErrCode := _iErrLatch;                                  // 故障期回放锁存码 / Replay the latched code during fault
ELSE
    iErrCode := _iInfoCode;                                  // 非故障期输出信息/降级码 / Info or degraded code outside fault
END_IF
IF _eState = E_DL_SPR_STATE.eIdle THEN
    sMsg := 'IDLE';                                          // 空闲 / Idle
ELSIF _eState = E_DL_SPR_STATE.eFeed THEN
    sMsg := 'FEED';                                          // 进泥 / Feeding
ELSIF _eState = E_DL_SPR_STATE.eMix THEN
    sMsg := 'MIX';                                           // 混合 / Mixing
ELSIF _eState = E_DL_SPR_STATE.ePress THEN
    sMsg := 'PRESS';                                         // 压榨 / Pressing
ELSIF _eState = E_DL_SPR_STATE.eFlush THEN
    sMsg := 'FLUSH';                                         // 冲洗 / Flushing
ELSIF _eState = E_DL_SPR_STATE.eRetract THEN
    sMsg := 'RETRACT';                                       // 退让 / Retracting
ELSE
    sMsg := 'FAULT';                                         // 故障 / Fault
END_IF
END_FUNCTION_BLOCK

(* ---- FB_DL_ScrubberReagentDoseSeq.st ---- *)
(*
  道莅工业代码库 / Daoli Industrial ST Library
  组件: FB_DL_ScrubberReagentDoseSeq
  分类: DL_Process
  复杂度: C4 ｜ 版本: 1.0.0 ｜ 2026-11-24
  平台兼容: CODESYS 3.5+ / TwinCAT 3 / 汇川 InoProShop / 施耐德 Machine Expert
  开源溯源: 无（clean-room 工程算法自研；参考公开的湿式洗涤塔 pH 反馈加碱与电导排污工艺，
            未复制任何受版权保护代码）
  许可证: 本项目自有 (MIT)

  功能职责:
    湿式洗涤塔碱液投加闭环。pH 反馈经简化 PI 调节计量泵，pH 稳定后进入保持态；
    循环液电导超限触发补排水（blowdown）；药剂罐低液位锁停计量泵并告警；
    泵运行中罐位下降率超限判泄漏疑似（安全侧）。

  输入/输出契约:
    IN  bEnable 上升沿启动（并做四项参数校验）；FALSE 撤销输出回 eIdle（R191 声明）。
    IN  bReset 上升沿是 eFault 唯一出口（还须残留故障条件消失）。
    OUT rPumpLh 计量泵冲程设定 [L/h]，仅在 eDose / eStabilize 输出，其余相为 0。
    OUT bMakeupValve / bDrainValve 仅在 eBlowdown 开，eFault 与 eTankLow 全关。

  码表 (Codes):
    31 = 药剂罐低液位（告警级；转 eTankLow，泵停，手动/上游补液）
    32 = 药液泄漏疑似（故障级；泵开时罐位下降率 > 5%/min）
    33 = 电导上限设定无效（故障级；rCondHi ≤ 0，比判据失效）
    34 = 计量泵上限无效（故障级；rPumpMaxLh ≤ 0，无饱和载体且增益不可算）
    35 = pH 测量值非法（故障级；越 0..14 或非有限）
    36 = 电导超限进入补排（信息级；blowdown 起点）
    37 = 补排次数达上限（故障级；反复补排说明补水/排污能力失效）
    38 = pH 设定值非法（故障级；rPhSp 越 0..14 或非有限）
    99 = 非法状态枚举值（ELSE 兜底）

  边界与红线:
    ① 五个定时器与两个 R_TRIG 全在 CASE 外无条件刷新（R7），CASE 内只读 .Q。
    ② tonStable / tonLow 的 IN 串本相或监测相闸并带 NOT .Q 自复位（R188）；tonLow 覆盖
       eDose/eStabilize/eBlowdown 三相，属**跨相累计看门狗**（低液位持续判定，与单相超时
       无关，红线 14 显式声明）；tonIntWin / tonDropWin 是自由运行周期窗（1 s 积分步 /
       60 s 下降率窗），不属任何相。
    ③ 积分 _rInteg 的显式清零条件：进 eIdle、进 eFault、进 eTankLow 三处即清（抗饱和载体
       同时把积分钳在 [0, rPumpMaxLh]）。
    ④ R528：bEnable 必须上升沿且泵上限/电导上限/pH 值/pH 设定四项有效才迁 eDose 或 eTankLow；
       全默认引脚时停留 eIdle，绝不直达投加相或补排相。
    ⑤ eFault 出口 = rtReset.Q AND NOT _bFaultCondNow（逐码反算残留条件，R28 可达性）。
    ⑥ 防抖硬性：电导补排出口用回差 DL_SCR_COND_HYST（禁零回差，否则在限值附近抖动会每拍
       进出补排相并迅速耗尽补排计数误报码 37）；泄漏判据 _bLeakNow 只在 60 s 窗边界采样一拍，
       禁把窗内旧差值当连续量逐拍复判（陈旧值复报会把一次骤降放大成永久故障）。
  修订历史: 2026-11-24  v1.0.0  R82-B 首版
*)

TYPE E_DL_SCRUB_STATE :
(
    eIdle      := 0,    // 空闲：等使能上升沿 / Idle: waiting for the enable rising edge
    eDose      := 1,    // 投加相：PI 调节计量泵 / Dose phase: PI control of the dosing pump
    eStabilize := 2,    // 稳定相：pH 在带内保持，等稳定确认 / Stabilize: pH inside the band, waiting for confirmation
    eBlowdown  := 3,    // 补排相：电导超限，开补水与排污阀 / Blowdown: conductivity high, makeup and drain valves open
    eTankLow   := 4,    // 低液位相：泵停告警，等罐位恢复 / Tank low: pump stopped with an alarm, waiting for recovery
    eFault     := 5     // 故障安全相：全部执行输出 FALSE / Fault safe phase: all actuator outputs FALSE
);
END_TYPE

FUNCTION_BLOCK FB_DL_ScrubberReagentDoseSeq
VAR_INPUT
    bEnable        : BOOL := FALSE;      // 使能（上升沿启动；FALSE 撤销输出回空闲）/ Enable, rising edge starts, FALSE withdraws the outputs
    bReset         : BOOL := FALSE;      // 复位（上升沿，eFault 唯一出口）/ Reset rising edge, the only fault exit
    rPh            : REAL := 0.0;        // 循环液 pH 实测 [-]/ Measured circulating liquid pH [-]
    rPhSp          : REAL := 0.0;        // pH 设定 [-]/ pH setpoint [-]
    rCondMsCm      : REAL := 0.0;        // 循环液电导率 [mS/cm] / Circulating liquid conductivity [mS/cm]
    rCondHi        : REAL := 0.0;        // 电导排污上限 [mS/cm] / Conductivity blowdown limit [mS/cm]
    rTankPct       : REAL := 0.0;        // 药剂罐余量 [%] / Reagent tank level [%]
    rTankLoPct     : REAL := 0.0;        // 药剂罐低液位阈值 [%] / Reagent tank low level threshold [%]
    rPumpMaxLh     : REAL := 0.0;        // 计量泵最大流量 [L/h] / Dosing pump maximum flow [L/h]
    tPhStable      : TIME := T#60S;      // pH 稳定确认时长，有效域 100ms..2h [s] / pH stability confirmation, valid domain 100ms..2h
    tTankLowDelay  : TIME := T#5S;       // 低液位确认时长，有效域 100ms..2h [s] / Low level confirmation, valid domain 100ms..2h
END_VAR
VAR_OUTPUT
    rPumpLh        : REAL := 0.0;        // 计量泵冲程设定 [L/h] / Dosing pump stroke setpoint [L/h]
    bPumpOn        : BOOL := FALSE;      // 计量泵运行位（单稳态，每拍重算）/ Pump run bit, monostable, recomputed every scan
    bMakeupValve   : BOOL := FALSE;      // 补水阀（仅补排相）/ Makeup valve, blowdown phase only
    bDrainValve    : BOOL := FALSE;      // 排污阀（仅补排相）/ Drain valve, blowdown phase only
    iErrCode       : INT := 0;           // 错误码（故障期锁存回放）/ Error code, latched replay during fault
    sMsg           : STRING;             // 文本提示（当前相位摘要）/ Text message, a summary of the current phase
END_VAR
VAR
    _eState        : E_DL_SCRUB_STATE := E_DL_SCRUB_STATE.eIdle;   // 内部相位（CASE 唯一写入目标）/ Internal phase, the only CASE write target
    _bFaultLatch   : BOOL := FALSE;      // 故障锁存位 / Fault latch
    _iErrLatch     : INT := 0;           // 锁存故障码（故障期唯一回放源）/ Latched fault code, the only replay source during fault
    _iInfoCode     : INT := 0;           // 信息级/告警级码 / Info or warning code
    _iErrTmp       : INT := 0;           // 当拍故障首因中间量 / First fault cause of this scan
    _bFaultReq     : BOOL := FALSE;      // 当拍故障请求（段 6 统一锁存）/ Fault request of this scan, latched at segment 6
    _bFaultCondNow : BOOL := FALSE;      // 残留故障条件（eFault 出口唯一附加判据）/ Residual fault condition, the only extra fault-exit criterion
    _bPhInvalid    : BOOL := FALSE;      // pH 测量值非法标志 / Measured pH invalid flag
    _bSpInvalid    : BOOL := FALSE;      // pH 设定值非法标志 / pH setpoint invalid flag
    _bStable       : BOOL := FALSE;      // 稳定确认记忆位（防 eDose↔eStabilize 每拍抖动）/ Stability memory, prevents scan-by-scan chatter
    _bLeakNow      : BOOL := FALSE;      // 泄漏疑似本拍成立（仅在 60 s 窗边界采样，防陈旧值复报）/ Leak suspicion valid in this scan, sampled only at the sixty second boundary
    _rPhCl         : REAL := 0.0;        // pH 净化副本 [-]/ Sanitised pH copy [-]
    _rSpCl         : REAL := 0.0;        // pH 设定净化副本 [-]/ Sanitised setpoint copy [-]
    _rCondCl       : REAL := 0.0;        // 电导率净化副本 [mS/cm] / Sanitised conductivity copy [mS/cm]
    _rCondExit     : REAL := 0.0;        // 补排出口门限（带回差，防抖）[mS/cm] / Blowdown exit threshold with hysteresis [mS/cm]
    _rTankCl       : REAL := 0.0;        // 罐位净化副本 [%] / Sanitised tank level copy [%]
    _rLoPct        : REAL := 0.0;        // 低液位阈值净化值 [%] / Sanitised low level threshold [%]
    _rErr          : REAL := 0.0;        // pH 误差 = 设定 - 实测 [pH] / pH error, setpoint minus measurement [pH]
    _rKp           : REAL := 0.0;        // 比例增益 [L/h per pH] / Proportional gain [L/h per pH]
    _rKi           : REAL := 0.0;        // 积分增益 [L/h per pH per s] / Integral gain [L/h per pH per s]
    _rIntMax       : REAL := 0.0;        // 积分上限（抗饱和载体）[L/h] / Integral upper limit, the anti-windup carrier [L/h]
    _rInteg        : REAL := 0.0;        // 积分项 [L/h] / Integral term [L/h]
    _rPumpCmd      : REAL := 0.0;        // 当拍泵设定 [L/h] / Pump command of this scan [L/h]
    _rPumpMax      : REAL := 0.0;        // 泵上限净化值 [L/h] / Sanitised pump maximum [L/h]
    _rDropPctMin   : REAL := 0.0;        // 罐位下降率（60 s 窗）[%/min] / Tank level drop rate over the sixty second window [%/min]
    _rTankPrevWin  : REAL := 0.0;        // 上一窗罐位快照 [%] / Tank level snapshot of the previous window [%]
    _iBlowdownCnt  : INT := 0;           // 补排次数，容量载体 DL_SCR_BD_MAX [次] / Blowdown counter, capacity carrier DL_SCR_BD_MAX [count]
    _tStable       : TIME := T#60S;      // pH 稳定确认钳定值 [s] / Clamped stability confirmation [s]
    _tLowDelay     : TIME := T#5S;       // 低液位确认钳定值 [s] / Clamped low level confirmation [s]
    rtReset        : R_TRIG;             // bReset 边沿（段 3 无条件刷新）/ bReset edge, refreshed unconditionally
    rtEnable       : R_TRIG;             // bEnable 边沿（段 3 无条件刷新，R528）/ bEnable edge, refreshed unconditionally
    tonStable      : TON;                // pH 稳定确认计时（本相单发，自复位）/ pH stability timer, single shot in its phase
    tonLow         : TON;                // 低液位累计看门狗（跨相持续判定，自复位）/ Low level cumulative watchdog across monitoring phases
    tonIntWin      : TON;                // 1 s 自由运行积分窗（自复位）/ One second free running integration window
    tonDropWin     : TON;                // 60 s 自由运行下降率窗（自复位）/ Sixty second free running drop rate window
END_VAR
VAR CONSTANT
    DL_SCR_EPS         : REAL := 1.0E-6;   // 数值闸阈值 [-]/ Numeric guard threshold [-]
    DL_SCR_FIN         : REAL := 1.0E15;   // 非有限判据阈值（ABS 比较用）[-] / Non-finite criterion threshold, compared by ABS [-]
    DL_SCR_PH_MIN      : REAL := 0.0;      // pH 有效域下限 [pH] / pH valid domain lower bound [pH]
    DL_SCR_PH_MAX      : REAL := 14.0;     // pH 有效域上限 [pH] / pH valid domain upper bound [pH]
    DL_SCR_PH_BAND     : REAL := 0.2;      // pH 稳定带宽 ±0.2 [pH] / pH stability band of plus or minus 0.2 [pH]
    DL_SCR_PH_SPAN     : REAL := 2.0;      // 比例增益折算满量程 pH 偏差 [pH] / pH deviation span used to scale the proportional gain [pH]
    DL_SCR_KI_RATIO    : REAL := 0.05;     // 积分增益 / 比例增益之比（每 1 s 步）[1/s] / Integral to proportional gain ratio per one second step [1/s]
    DL_SCR_INT_RATIO   : REAL := 1.0;      // 积分上限 / 泵上限之比 [-] / Integral limit to pump maximum ratio [-]
    DL_SCR_TANK_HYST   : REAL := 5.0;      // 低液位恢复回差 [%] / Low level recovery hysteresis [%]
    DL_SCR_DROP_LIM    : REAL := 5.0;      // 罐位下降率泄漏阈值 [%/min] / Tank drop rate leak threshold [%/min]
    DL_SCR_COND_HYST   : REAL := 0.5;      // 电导补排回差（防抖，禁零回差）[mS/cm] / Conductivity blowdown hysteresis, chatter prevention [mS/cm]
    DL_SCR_BD_MAX      : INT := 6;         // 单使能周期补排次数上限 [次] / Blowdown count limit per enable cycle [count]
    DL_SCR_ONE         : INT := 1;         // 计数步进一 [1] / Counter step of one [1]
    DL_SCR_ZERO        : INT := 0;         // 计数零基准 [-] / Counter zero base [-]
    DL_SCR_T_MIN       : TIME := T#100MS;  // 时间参数下限 [s] / Time parameter lower bound [s]
    DL_SCR_T_MAX       : TIME := T#2H;     // 时间参数上限 [s] / Time parameter upper bound [s]
    DL_SCR_T_STABLE_DEF: TIME := T#60S;    // 稳定确认默认回退值（在域内）[s] / Default stability duration inside the domain [s]
    DL_SCR_T_LOW_DEF   : TIME := T#5S;     // 低液位确认默认回退值（在域内）[s] / Default low level duration inside the domain [s]
    DL_SCR_INTWIN      : TIME := T#1S;     // 积分步长窗 [s] / Integration step window [s]
    DL_SCR_DROPWIN     : TIME := T#60S;    // 下降率测量窗 [s] / Drop rate measurement window [s]
END_VAR

(* —— 段 1：中间量预置（只清当拍扫描量，不清锁存/积分/补排计数，FB32-1） —— *)
_iErrTmp   := 0;                                    // 当拍故障首因复位 / Scan first fault cause reset
_bFaultReq := FALSE;                                // 当拍故障请求复位 / Scan fault request reset

(* —— 段 2：时间参数两级回退 + 入参域闸与非有限兜底 + 增益折算 —— *)
IF (tPhStable < DL_SCR_T_MIN) OR (tPhStable > DL_SCR_T_MAX) THEN
    _tStable := DL_SCR_T_STABLE_DEF;                // 越域：回一级默认常量 / Out of domain: fall back to the default constant
ELSE
    _tStable := tPhStable;                          // 域内：原值采用 / Inside the domain: use as given
END_IF
IF (tTankLowDelay < DL_SCR_T_MIN) OR (tTankLowDelay > DL_SCR_T_MAX) THEN
    _tLowDelay := DL_SCR_T_LOW_DEF;                 // 越域：回一级默认常量 / Out of domain: fall back to the default constant
ELSE
    _tLowDelay := tTankLowDelay;                    // 域内：原值采用 / Inside the domain: use as given
END_IF
_bPhInvalid := FALSE;                               // pH 非法标志预置 / Invalid pH flag preset
_rPhCl      := rPh;                                 // pH 副本 [-]/ pH copy [-]
IF (ABS(_rPhCl) > DL_SCR_FIN) OR (_rPhCl < DL_SCR_PH_MIN) OR (_rPhCl > DL_SCR_PH_MAX) THEN
    _bPhInvalid := TRUE;                            // 非有限或越 0..14：参与判据前必须先拦 / Non-finite or out of zero to fourteen: block it before it feeds any criterion
    _rPhCl      := DL_SCR_PH_MIN;                   // 兜底钳到域下限（值不参与结论）/ Clamp to the lower bound, the value never feeds a decision
END_IF
_bSpInvalid := FALSE;                               // 设定非法标志预置 / Invalid setpoint flag preset
_rSpCl      := rPhSp;                               // 设定副本 [-]/ Setpoint copy [-]
IF (ABS(_rSpCl) > DL_SCR_FIN) OR (_rSpCl < DL_SCR_PH_MIN) OR (_rSpCl > DL_SCR_PH_MAX) THEN
    _bSpInvalid := TRUE;                            // 非有限或越 0..14 / Non-finite or out of zero to fourteen
    _rSpCl      := DL_SCR_PH_MIN;                   // 兜底钳到域下限（值不参与结论）/ Clamp to the lower bound, the value never feeds a decision
END_IF
_rCondCl := rCondMsCm;                              // 电导率副本 [mS/cm] / Conductivity copy [mS/cm]
IF (ABS(_rCondCl) > DL_SCR_FIN) OR (_rCondCl < 0.0) THEN
    _rCondCl := 0.0;                                // 非有限或负值兜底为零 / Non-finite or negative falls back to zero
END_IF
_rCondExit := rCondHi - DL_SCR_COND_HYST;           // 量纲: (mS/cm)-(mS/cm) = mS/cm 补排出口门限 / Blowdown exit threshold in mS/cm
IF (ABS(rCondHi) > DL_SCR_FIN) OR (_rCondExit < 0.0) THEN
    _rCondExit := 0.0;                              // 非有限或负门限兜底为零（保证出口可达）/ Non-finite or negative falls back to zero so the exit stays reachable
END_IF
_rTankCl := rTankPct;                               // 罐位副本 [%] / Tank level copy [%]
IF (ABS(_rTankCl) > DL_SCR_FIN) OR (_rTankCl < 0.0) THEN
    _rTankCl := 0.0;                                // 非有限或负值兜底为零 / Non-finite or negative falls back to zero
ELSIF _rTankCl > 100.0 THEN
    _rTankCl := 100.0;                              // 罐位上限饱和 [%] / Saturate the tank level at one hundred percent
END_IF
_rLoPct := rTankLoPct;                              // 低液位阈值副本 [%] / Low level threshold copy [%]
IF (ABS(_rLoPct) > DL_SCR_FIN) OR (_rLoPct < 0.0) THEN
    _rLoPct := 0.0;                                 // 非有限或负值兜底为零 / Non-finite or negative falls back to zero
ELSIF _rLoPct > 95.0 THEN
    _rLoPct := 95.0;                                // 阈值上限饱和，保证恢复回差可达 [%] / Saturate so the recovery hysteresis stays reachable [%]
END_IF
_rPumpMax := rPumpMaxLh;                            // 泵上限副本 [L/h] / Pump maximum copy [L/h]
IF (ABS(_rPumpMax) > DL_SCR_FIN) OR (_rPumpMax < 0.0) THEN
    _rPumpMax := 0.0;                               // 非有限或负值兜底为零 / Non-finite or negative falls back to zero
END_IF
_rErr := _rSpCl - _rPhCl;                           // 误差取「设定减实测」：pH 低于设定为正 → 泵加量（碱液）/ Error is setpoint minus measurement, a low pH gives a positive dose
IF _rPumpMax > DL_SCR_EPS THEN
    _rKp     := _rPumpMax / DL_SCR_PH_SPAN;         // 量纲: (L/h)/(pH) = L/h per pH / (L/h) divided by (pH) gives L/h per pH
    _rKi     := _rKp * DL_SCR_KI_RATIO;             // 量纲: (L/h per pH)*(1/s) = L/h per pH per s / (L/h per pH) times (1/s)
    _rIntMax := _rPumpMax * DL_SCR_INT_RATIO;       // 量纲: (L/h)*(无量纲) = L/h（积分上限载体）/ (L/h) times dimensionless gives the integral carrier
ELSE
    _rKp     := 0.0;                                // 分母闸：泵上限无效时增益置零 / Denominator guard: gains are zero when the pump limit is invalid
    _rKi     := 0.0;                                // 分母闸：积分增益置零 / Denominator guard: the integral gain is zero
    _rIntMax := 0.0;                                // 分母闸：积分上限置零 / Denominator guard: the integral limit is zero
END_IF
_bFaultCondNow := FALSE;                            // 残留条件预置（eFault 出口唯一附加判据）/ Residual preset, the only extra fault-exit criterion
IF _iErrLatch = 33 THEN
    _bFaultCondNow := (ABS(rCondHi) <= DL_SCR_EPS);         // 码 33：电导上限仍无效 / Code 33: the conductivity limit is still invalid
ELSIF _iErrLatch = 34 THEN
    _bFaultCondNow := (rPumpMaxLh <= DL_SCR_EPS);           // 码 34：泵上限仍无效 / Code 34: the pump limit is still invalid
ELSIF _iErrLatch = 35 THEN
    _bFaultCondNow := _bPhInvalid;                          // 码 35：pH 测量仍非法 / Code 35: the measured pH is still invalid
ELSIF _iErrLatch = 38 THEN
    _bFaultCondNow := _bSpInvalid;                          // 码 38：pH 设定仍非法 / Code 38: the pH setpoint is still invalid
END_IF
(* 码 32（泄漏疑似）以「泵运行中的下降率」为必要条件，故障相泵已停、条件自然不再成立；
   码 37（补排次数达上限）由计数驱动。二者与码 99 均无输入残留条件，复位沿单独即可退出。 / Codes 32, 37 and 99 have no residual input condition *)

(* —— 段 3：边沿与定时器（全部在 CASE 外无条件刷新，R7；IN 带 NOT .Q 自复位，R188） —— *)
rtReset(CLK := bReset);                             // 复位边沿无条件刷新 / Reset edge refreshed unconditionally
rtEnable(CLK := bEnable);                           // 使能边沿无条件刷新（R528 起点判据）/ Enable edge refreshed unconditionally
tonStable(IN := (_eState = E_DL_SCRUB_STATE.eStabilize) AND (NOT tonStable.Q) AND (NOT _bFaultLatch),
          PT := _tStable);                          // 本相单发计时：仅稳定相 / Single-shot timer in the stabilize phase only
tonLow(IN := ((_eState = E_DL_SCRUB_STATE.eDose) OR (_eState = E_DL_SCRUB_STATE.eStabilize)
              OR (_eState = E_DL_SCRUB_STATE.eBlowdown))
             AND (_rTankCl <= _rLoPct) AND (NOT tonLow.Q) AND (NOT _bFaultLatch),
       PT := _tLowDelay);                           // 跨相累计看门狗：低液位在三监测相内持续累计，非本相超时 / Cumulative watchdog across the three monitoring phases, not a phase timeout
tonIntWin(IN := NOT tonIntWin.Q, PT := DL_SCR_INTWIN);      // 自由运行 1 s 积分步长窗 / Free running one second integration step window
tonDropWin(IN := NOT tonDropWin.Q, PT := DL_SCR_DROPWIN);   // 自由运行 60 s 下降率测量窗 / Free running sixty second drop rate window
IF tonIntWin.Q THEN
    IF (_eState = E_DL_SCRUB_STATE.eDose) AND (NOT _bFaultLatch) THEN
        // 量纲: (pH)*(L/h per pH per s)*(1 s) = L/h 积分增量（窗长即 1 s，故不再乘 dt）
        _rInteg := _rInteg + (_rErr * _rKi);        // 积分项一步累加 [L/h] / One integration step [L/h]
        IF _rInteg > _rIntMax THEN
            _rInteg := _rIntMax;                    // 抗饱和上限 / Anti-windup upper clamp
        END_IF
        IF _rInteg < 0.0 THEN
            _rInteg := 0.0;                         // 抗饱和下限 / Anti-windup lower clamp
        END_IF
    END_IF
END_IF
IF tonDropWin.Q THEN
    // 量纲: (% 窗内差) / (60 s 窗) * 60 s = %/min；窗长已是 60 s，故差值即 %/min
    _rDropPctMin  := _rTankPrevWin - _rTankCl;      // 窗内罐位下降百分点 [%/min] / Tank drop in percentage points over the window [%/min]
    _rTankPrevWin := _rTankCl;                      // 刷新下一窗快照 [%] / Refresh the snapshot for the next window [%]
END_IF

(* —— 段 4：当拍泵设定（PI 简化：pump = kp*err + integ，限幅 [0, rPumpMaxLh]） —— *)
IF _rPumpMax > DL_SCR_EPS THEN
    // 量纲: (L/h per pH)*(pH) + (L/h) = L/h
    _rPumpCmd := (_rKp * _rErr) + _rInteg;          // PI 输出 [L/h] / PI output [L/h]
    IF _rPumpCmd > _rPumpMax THEN
        _rPumpCmd := _rPumpMax;                     // 上限饱和（载体 rPumpMaxLh）/ Saturate at the pump maximum
    END_IF
    IF _rPumpCmd < 0.0 THEN
        _rPumpCmd := 0.0;                           // 下限饱和，禁负投加 / Saturate at zero, no negative dosing
    END_IF
ELSE
    _rPumpCmd := 0.0;                               // 分母闸：泵上限无效则出零 / Denominator guard: emit zero when the pump limit is invalid
END_IF
_bLeakNow := FALSE;                                 // 泄漏判据预置 / Leak criterion preset
IF tonDropWin.Q AND (_rDropPctMin > DL_SCR_DROP_LIM) AND (_rPumpCmd > DL_SCR_EPS)
   AND ((_eState = E_DL_SCRUB_STATE.eDose) OR (_eState = E_DL_SCRUB_STATE.eStabilize)) THEN
    _bLeakNow := TRUE;                              // 窗边界单拍采样：泵在开且窗内罐位骤降，泄漏疑似 / Sampled once per window boundary
END_IF

(* —— 段 5：状态机主体（唯一相位写入点；故障只置请求，锁存与迁相由段 6 执行） —— *)
CASE _eState OF
    E_DL_SCRUB_STATE.eIdle :
        (* 迁移①：拍 N 进入（使能上升沿）/ 本拍行为：四项参数校验，缺任一即故障 / 拍 N+1 转出至投加相或低液位相 *)
        IF rtEnable.Q AND (NOT _bFaultLatch) THEN
            IF rPumpMaxLh <= DL_SCR_EPS THEN
                _iErrTmp   := 34;                            // 故障级：泵上限无效 / Fault: invalid pump maximum
                _bFaultReq := TRUE;                          // 请求段 6 锁存 / Request the latch at segment 6
            ELSIF ABS(rCondHi) <= DL_SCR_EPS THEN
                _iErrTmp   := 33;                            // 故障级：电导上限无效 / Fault: invalid conductivity limit
                _bFaultReq := TRUE;                          // 请求段 6 锁存 / Request the latch at segment 6
            ELSIF _bPhInvalid THEN
                _iErrTmp   := 35;                            // 故障级：pH 测量非法 / Fault: invalid pH measurement
                _bFaultReq := TRUE;                          // 请求段 6 锁存 / Request the latch at segment 6
            ELSIF _bSpInvalid THEN
                _iErrTmp   := 38;                            // 故障级：pH 设定非法 / Fault: invalid pH setpoint
                _bFaultReq := TRUE;                          // 请求段 6 锁存 / Request the latch at segment 6
            ELSIF _rTankCl <= _rLoPct THEN
                _rInteg        := 0.0;                       // 进低液位相即清积分 / Integral cleared on entry to the low level phase
                _iBlowdownCnt  := DL_SCR_ZERO;               // 新周期补排计数归零 / New cycle: blowdown counter cleared
                _iInfoCode     := 31;                        // 告警级：起始即低液位 / Warning: low level at start
                _eState        := E_DL_SCRUB_STATE.eTankLow;  // 迁移①：进低液位相 / Move to the tank low phase
            ELSE
                _rInteg        := 0.0;                       // 新周期：清积分 / New cycle: integral cleared
                _iBlowdownCnt  := DL_SCR_ZERO;               // 新周期：补排计数归零 / New cycle: blowdown counter cleared
                _bStable       := FALSE;                     // 新周期：稳定记忆清零 / New cycle: stability memory cleared
                _iInfoCode     := 0;                         // 新周期：信息码归零 / New cycle: info code cleared
                _eState        := E_DL_SCRUB_STATE.eDose;    // 迁移①：进投加相 / Move to the dose phase
            END_IF
        END_IF

    E_DL_SCRUB_STATE.eDose :
        (* 迁移②③④：拍 N 进入 / 本拍行为：PI 输出泵设定；逐拍查低液位、电导超限 / 拍 N+1 转出 *)
        IF tonLow.Q THEN                                         // 低液位经 tTankLowDelay 确认（累计看门狗）才锁停 / Locked out only after the delay confirms
            _rInteg    := 0.0;                               // 进低液位相即清积分 / Integral cleared on entry
            _iInfoCode := 31;                                // 告警级：低液位 / Warning: low level
            _eState    := E_DL_SCRUB_STATE.eTankLow;         // 迁移②：锁停计量泵 / Stop the dosing pump
        ELSIF _rCondCl > rCondHi THEN
            _iInfoCode := 36;                                // 信息级：电导超限进补排 / Info: conductivity high, entering blowdown
            IF _iBlowdownCnt < DL_SCR_BD_MAX THEN
                _iBlowdownCnt := _iBlowdownCnt + DL_SCR_ONE; // 补排次数净额 +1，达容量上限饱和 / Net blowdown increment, saturated at capacity
            END_IF
            IF _iBlowdownCnt >= DL_SCR_BD_MAX THEN
                _iErrTmp   := 37;                            // 故障级：反复补排说明补水/排污失效 / Fault: repeated blowdown means makeup or drain has failed
                _bFaultReq := TRUE;                          // 请求段 6 锁存 / Request the latch at segment 6
            ELSE
                _eState := E_DL_SCRUB_STATE.eBlowdown;       // 迁移③：进补排相 / Move to blowdown
            END_IF
        ELSIF (ABS(_rErr) <= DL_SCR_PH_BAND) AND (NOT _bStable) THEN
            _eState := E_DL_SCRUB_STATE.eStabilize;          // 迁移④：进带内，转稳定确认相 / In band, move to the stabilize phase
        ELSE
            IF ABS(_rErr) > DL_SCR_PH_BAND THEN
                _bStable := FALSE;                           // 出带即撤销稳定确认 / Leaving the band revokes the stability memory
            END_IF
        END_IF

    E_DL_SCRUB_STATE.eStabilize :
        (* 迁移⑤⑥⑦：拍 N 进入 / 本拍行为：pH 保持在带内才计稳定；出带回投加相 / 拍 N+1 转出 *)
        IF tonLow.Q THEN                                         // 低液位经 tTankLowDelay 确认（累计看门狗）才锁停 / Locked out only after the delay confirms
            _rInteg    := 0.0;                               // 进低液位相即清积分 / Integral cleared on entry
            _iInfoCode := 31;                                // 告警级：低液位 / Warning: low level
            _eState    := E_DL_SCRUB_STATE.eTankLow;         // 迁移⑤：锁停计量泵 / Stop the dosing pump
        ELSIF _rCondCl > rCondHi THEN
            _iInfoCode := 36;                                // 信息级：电导超限进补排 / Info: conductivity high, entering blowdown
            IF _iBlowdownCnt < DL_SCR_BD_MAX THEN
                _iBlowdownCnt := _iBlowdownCnt + DL_SCR_ONE; // 补排次数净额 +1 / Net blowdown increment
            END_IF
            IF _iBlowdownCnt >= DL_SCR_BD_MAX THEN
                _iErrTmp   := 37;                            // 故障级：补排次数达上限 / Fault: blowdown count at its limit
                _bFaultReq := TRUE;                          // 请求段 6 锁存 / Request the latch at segment 6
            ELSE
                _eState := E_DL_SCRUB_STATE.eBlowdown;       // 迁移⑥：进补排相 / Move to blowdown
            END_IF
        ELSIF ABS(_rErr) > DL_SCR_PH_BAND THEN
            _bStable := FALSE;                               // 出带：撤销稳定确认 / Left the band: revoke the stability memory
            _eState  := E_DL_SCRUB_STATE.eDose;              // 迁移⑦：回投加相继续调节 / Back to dose and keep regulating
        ELSIF tonStable.Q THEN
            _bStable   := TRUE;                              // 稳定确认成立（保持态）/ Stability confirmed, hold state
            _iInfoCode := 0;                                 // 稳定达成：清信息码 / Stable: info code cleared
            _eState    := E_DL_SCRUB_STATE.eDose;            // 迁移⑦：回投加相保持 / Back to dose in the hold state
        END_IF

    E_DL_SCRUB_STATE.eBlowdown :
        (* 迁移⑧⑨：拍 N 进入 / 本拍行为：开补水与排污，泵停 / 拍 N+1 转出至投加相或低液位相 *)
        IF tonLow.Q THEN                                         // 低液位经 tTankLowDelay 确认（累计看门狗）才锁停 / Locked out only after the delay confirms
            _rInteg    := 0.0;                               // 进低液位相即清积分 / Integral cleared on entry
            _iInfoCode := 31;                                // 告警级：低液位 / Warning: low level
            _eState    := E_DL_SCRUB_STATE.eTankLow;         // 迁移⑧：补排中低液位，锁停 / Low level during blowdown, stop
        ELSIF _rCondCl < _rCondExit THEN
            _bStable := FALSE;                               // 补排结束：撤销稳定确认 / Blowdown done: revoke the stability memory
            _eState  := E_DL_SCRUB_STATE.eDose;              // 迁移⑨：电导回落到回差下，回投加相 / Conductivity fell below the hysteresis band, back to dose
        END_IF

    E_DL_SCRUB_STATE.eTankLow :
        (* 迁移⑩：拍 N 进入 / 本拍行为：泵停告警，等罐位回到 lo + 5% / 拍 N+1 转出至投加相 *)
        IF _rTankCl > (_rLoPct + DL_SCR_TANK_HYST) THEN
            _bStable   := FALSE;                             // 恢复补液：稳定需重新确认 / After refilling the stability must be re-confirmed
            _iInfoCode := 0;                                 // 恢复：清信息码 / Recovered: info code cleared
            _eState    := E_DL_SCRUB_STATE.eDose;            // 迁移⑩：回投加相 / Back to the dose phase
        END_IF

    E_DL_SCRUB_STATE.eFault :
        (* 迁移⑪：拍 N 进入 / 本拍行为：只等出口条件（复位沿 + 残留条件消失）/ 拍 N+1 转出至 eIdle *)
        IF rtReset.Q AND (NOT _bFaultCondNow) THEN
            _bFaultLatch  := FALSE;                          // 清故障锁存 / Clear the fault latch
            _iErrLatch    := 0;                              // 清锁存故障码 / Clear the latched code
            _iInfoCode    := 0;                              // 清信息码 / Clear the info code
            _rInteg       := 0.0;                            // 进 eIdle 前的积分清零 / Integral cleared before returning to idle
            _bStable      := FALSE;                          // 稳定记忆清零 / Stability memory cleared
            _iBlowdownCnt := DL_SCR_ZERO;                    // 补排计数清零 / Blowdown counter cleared
            _eState       := E_DL_SCRUB_STATE.eIdle;         // 回空闲相，不滞留 / Back to idle, never parked
        END_IF
ELSE
    (* 迁移⑫：非法枚举兜底（R6），码位赋值与锁存 3 行内配对（R45） *)
    IF NOT _bFaultLatch THEN
        _iErrLatch   := 99;                                  // 故障级：非法状态枚举值 / Fault: illegal state enum value
        _bFaultLatch := TRUE;                                // 置故障锁存 / Latch the fault
    END_IF
END_CASE

(* —— 段 6：泄漏疑似判定 + 故障锁存 + 段尾迁相 + 撤使能降级（R191 已声明） —— *)
IF _bLeakNow AND (NOT _bFaultLatch) THEN
    _iErrTmp   := 32;                                    // 故障级：泵运行中罐位骤降，泄漏疑似 / Fault: the tank level drops while pumping, a leak is suspected
    _bFaultReq := TRUE;                                  // 请求本次锁存 / Request the latch in this scan
END_IF
IF _bFaultReq AND (NOT _bFaultLatch) THEN
    _iErrLatch   := _iErrTmp;                            // 锁存当拍首因 / Latch the first cause of this scan
    _bFaultLatch := TRUE;                                // 置故障锁存 / Latch the fault
END_IF
IF _bFaultLatch AND (_eState <> E_DL_SCRUB_STATE.eFault) THEN
    _eState := E_DL_SCRUB_STATE.eFault;                  // 锁存即迁相（段尾统一执行）/ The latch forces the fault phase at the tail
END_IF
IF (NOT bEnable) AND (NOT _bFaultLatch) AND (_eState <> E_DL_SCRUB_STATE.eIdle) THEN
    _rInteg := 0.0;                                      // 撤使能：清积分（进 eIdle 条件之一）/ Disable: integral cleared
    _bStable := FALSE;                                   // 撤使能：清稳定记忆 / Disable: stability memory cleared
    _eState := E_DL_SCRUB_STATE.eIdle;                   // 撤使能：回空闲相 / Disable: back to idle
END_IF

(* —— 段 7：统一出口（单稳态每拍重算，不锁存；eFault 内全部 FALSE） —— *)
IF ((_eState = E_DL_SCRUB_STATE.eDose) OR (_eState = E_DL_SCRUB_STATE.eStabilize)) AND (NOT _bFaultLatch) THEN
    rPumpLh  := _rPumpCmd;                               // 投加相与稳定相输出泵设定 [L/h] / Dose and stabilize phases emit the pump setpoint [L/h]
    bPumpOn  := (_rPumpCmd > DL_SCR_EPS);                // 设定为正直才置运行位 / The run bit is set only for a positive setpoint
ELSE
    rPumpLh  := 0.0;                                     // 其余相（含补排、低液位、故障）：泵设定归零 / Other phases, including blowdown, low level and fault, emit zero
    bPumpOn  := FALSE;                                   // 其余相：运行位撤销 / Other phases: the run bit is withdrawn
END_IF
bMakeupValve := (_eState = E_DL_SCRUB_STATE.eBlowdown) AND (NOT _bFaultLatch);   // 补水阀仅补排相 / Makeup valve only during blowdown
bDrainValve  := (_eState = E_DL_SCRUB_STATE.eBlowdown) AND (NOT _bFaultLatch);   // 排污阀仅补排相 / Drain valve only during blowdown
IF _bFaultLatch THEN
    iErrCode := _iErrLatch;                              // 故障期回放锁存码 / Replay the latched code during fault
ELSE
    iErrCode := _iInfoCode;                              // 非故障期输出信息/告警码 / Info or warning code outside fault
END_IF
IF _eState = E_DL_SCRUB_STATE.eIdle THEN
    sMsg := 'IDLE';                                      // 空闲 / Idle
ELSIF _eState = E_DL_SCRUB_STATE.eDose THEN
    sMsg := 'DOSE';                                      // 投加 / Dosing
ELSIF _eState = E_DL_SCRUB_STATE.eStabilize THEN
    sMsg := 'STABLE';                                    // 稳定确认 / Stabilizing
ELSIF _eState = E_DL_SCRUB_STATE.eBlowdown THEN
    sMsg := 'BLOWDOWN';                                  // 补排 / Blowdown
ELSIF _eState = E_DL_SCRUB_STATE.eTankLow THEN
    sMsg := 'TANKLOW';                                   // 药罐低液位 / Reagent tank low
ELSE
    sMsg := 'FAULT';                                     // 故障 / Fault
END_IF
END_FUNCTION_BLOCK

(* ---- FB_DL_SealJawDwellTrim.st ---- *)
(*==============================================================================
 * 组件名称 (Component)  : FB_DL_SealJawDwellTrim
 * 所属子库 (Sublibrary) : DL_Process
 * 当前版本 (Version)    : 1.0.0
 * 兼容性 (Platform)     : CODESYS 3.5 / TwinCAT 3 / 汇川 InoProShop（纯标准元素，无方言）
 * 功能描述 (Function)   : 热封刀驻留时间随线速自整定（限速微调）。以封口质量对目标的偏差
 *                         按微调增益积分出驻留补偿量，先按变化率限速、再按上下限钳制
 *                         （反序会让爬升把超限带出来），停机期不计数、不积分；质量读数非
 *                         有限则冻结微调并保持上次给定（不把 NaN 积分进给定）。不做温控、
 *                         不做封口质量判定本身（由引脚注入）、不做多刀头协调。
 *                         遗留假设（代理阈值三句）：① 代理任务周期取 100 ms（本件无周期
 *                         引脚）；② 覆盖 50~200 ms 的任务周期，偏差 ≤2 倍；③ 更快的任务
 *                         周期由调用方在 fDwellRateMax_msS 上折算，本件不负责。
 * 溯源 (Origin)         : 道莅 clean-room 防御性实现
 * 本文件内含 (Contains) : TYPE E_DL_DwellState / FUNCTION_BLOCK FB_DL_SealJawDwellTrim
 * 依赖 (Depends)        : 无（仅 Standard.library 的 ABS / LIMIT / MIN / MAX）
 * 红线自检 (Redline)    : 无外部全局变量、无硬件地址直引 ｜ 全变量中英双语同行注释
 *                         上下限与目标判零防除零 ｜ 质量非有限即冻结微调并保持给定 ｜ 先限速
 *                         后钳制 ｜ 枚举显式赋值 ｜ CASE 含 ELSE 兜底 ｜ 本件无定时器/沿实例，
 *                         全部逻辑为无状态算术，故无周期刷新项
 * 错误码表 (Codes)      : 16#0005_043A 就绪（微调正常或停机冻结）
 *                         16#0005_043B 预留：本版不发码（下一轮区间起点，禁止回填）
 *                         16#0005_043C 故障级 组态非法（上下限反置、目标/增益/变化率出域）
 *                         16#0005_043D 信息级 驻留给定触限并已钳制（不置故障级标志）
 *                         16#0005_043E 故障级 质量读数非有限，微调冻结并保持上次给定
 * 修订历史 (Revision)   : 2026-11-17  v1.0.0  首版入库 · R28 · 阶段三批 4
 * 验收向量 (Acceptance) : 正向 标称 300 ms、线速 0→60 m/min、质量 0.85 对目标 0.90 → 微调
 *                         +10 ms、给定 310 ms、斜率 ≤50 ms/s
 *                         反向 下限设 400 ms > 上限 300 ms → 16#0005_043C；质量给 NaN →
 *                         16#0005_043E 且给定保持；给定顶到上限 → 16#0005_043D 且 bAtLimit
 *============================================================================*)

(*-----------------------------------------------------------------------------
 * 枚举: E_DL_DwellState（归属本功能块，同文件发布，全库唯一定义）
 *----------------------------------------------------------------------------*)
TYPE E_DL_DwellState :
(
    eFrozen  := 0,    // 冻结：停机、禁用或质量不可信 / Frozen, stopped, disabled or the quality is untrustworthy
    eTrim    := 10,   // 微调：限速 + 钳制后的驻留给定 / Trimming, rate limited and clamped
    eAtLimit := 20,   // 触限：给定顶在上下限 / At a limit, the setpoint sits on a bound
    eFault   := 99    // 故障：组态非法锁存 / Fault, the configuration error is latched
);
END_TYPE

FUNCTION_BLOCK FB_DL_SealJawDwellTrim
VAR_INPUT
    bEnable         : BOOL := FALSE;      // 使能 / Enable
    bRunning        : BOOL := FALSE;      // 线运行（停机冻结自整定） / Line running, tuning is frozen when stopped
    fLineSpeed_mpm  : REAL := 0.0;        // 线速度 [m/min]，域 0~200 / Line speed in metres per minute, domain 0 to 200
    fDwellNominal_ms : REAL := 300.0;     // 标称驻留 [ms]，域 50~2000 / Nominal dwell, domain 50 to 2000 ms
    fDwellMin_ms    : REAL := 200.0;      // 驻留下限 [ms] / Dwell lower bound
    fDwellMax_ms    : REAL := 500.0;      // 驻留上限 [ms]，须 > 下限 / Dwell upper bound, must exceed the lower bound
    fSealQuality    : REAL := 0.9;        // 封口质量 [0~1]（注入） / Seal quality from zero to one, injected
    fQualityTarget  : REAL := 0.9;        // 目标质量 [—]，域 0.7~0.99 / Quality target, domain 0.7 to 0.99
    fTrimGain       : REAL := 20.0;       // 微调增益 [ms/单位误差]，域 0~50 / Trim gain in milliseconds per unit error
    fDwellRateMax_msS : REAL := 50.0;     // 变化率上限 [ms/s]，域 1~200 / Rate limit in milliseconds per second
END_VAR
VAR_OUTPUT
    fDwellOut_ms    : REAL;               // 驻留给定 [ms] / Dwell setpoint in milliseconds
    fDwellTrim_ms   : REAL;               // 微调分量 [ms] / Trim component in milliseconds
    bAtLimit        : BOOL;               // 到上下限 / At a bound
    uTrimCnt        : UDINT;              // 微调生效次数 [次] / Effective trim count
    eErr            : UDINT;               // 错误码，段位 16#0005_xxxx / Error code in segment 16#0005_xxxx
END_VAR
VAR
    _eState         : E_DL_DwellState := E_DL_DwellState.eFrozen; // 当前相位 / Current phase
    _bInit          : BOOL := FALSE;      // 首扫标志，取非判定 / First-scan flag, tested negated
    _bCfgOk         : BOOL;               // 组态合法标志 / Configuration valid flag
    _bFaultLatch    : BOOL := FALSE;      // 组态故障锁存 / Configuration fault latch
    _bQualityOk     : BOOL;               // 质量读数可信标志 / Quality reading trustworthy flag
    _fErr           : REAL;               // 质量误差（目标 − 实测） / Quality error, target minus measured
    _fTrimWant      : REAL := 0.0;        // 期望微调分量 [ms] / Desired trim component
    _fTrimStep      : REAL;               // 本拍允许的微调步长 [ms] / Allowed trim step of this scan
    _fTrimDelta     : REAL;               // 本拍实际微调增量 [ms] / Actual trim increment of this scan
    _fDwellRaw      : REAL;               // 限速后驻留 [ms] / Rate-limited dwell
    _fDwellPrev     : REAL := 300.0;      // 上一拍驻留给定 [ms] / Previous dwell setpoint
END_VAR
VAR CONSTANT
    DL_DW_READY    : UDINT := 16#0005_043A;  // 就绪码 / Ready code
    DL_DW_CFG_BAD  : UDINT := 16#0005_043C;  // 故障级组态非法码 / Fault code for bad configuration
    DL_DW_LIMIT    : UDINT := 16#0005_043D;  // 信息级触限钳制码 / Info code for bound clamping
    DL_DW_QUAL_BAD : UDINT := 16#0005_043E;  // 故障级质量非有限码 / Fault code for a non-finite quality
    DL_DW_NOM_LO   : REAL := 50.0;           // 标称驻留下限 [ms] / Nominal dwell lower bound
    DL_DW_NOM_HI   : REAL := 2000.0;         // 标称驻留上限 [ms] / Nominal dwell upper bound
    DL_DW_TGT_LO   : REAL := 0.7;            // 目标质量下限 / Quality target lower bound
    DL_DW_TGT_HI   : REAL := 0.99;           // 目标质量上限 / Quality target upper bound
    DL_DW_GAIN_HI  : REAL := 50.0;           // 增益上限 [ms/单位误差] / Gain upper bound
    DL_DW_RATE_LO  : REAL := 1.0;            // 变化率下限 [ms/s] / Rate lower bound
    DL_DW_RATE_HI  : REAL := 200.0;          // 变化率上限 [ms/s] / Rate upper bound
    DL_DW_TASK_S   : REAL := 0.1;            // 代理任务周期 [s]（遗留假设） / Proxy task period in seconds
    DL_DW_TRIM_EPS : REAL := 1.0;            // 微调计数门限 [ms] / Trim counting threshold
END_VAR

// 段 1｜输出与单拍标志预置
bAtLimit := FALSE;                                  // 触限标志预清 / At-bound flag pre-cleared
eErr := 0;                                          // 错误码预清 / Error code pre-cleared

// 段 2｜首扫初始化（判据取非，R19）
IF NOT _bInit THEN
    _fTrimWant := 0.0;                              // 微调起点 0 [ms] / Trim starts at zero
    _fDwellPrev := fDwellNominal_ms;                // 上一拍驻留取标称 [ms] / Previous dwell starts from the nominal value
    _eState := E_DL_DwellState.eFrozen;             // 相位冻结起步 / Phase starts frozen
    _bInit := TRUE;                                 // 首扫只做一次 / The first scan runs once
END_IF

// 段 3｜组态闸（上下限反置 → 微调区间为空；目标与变化率出域）
_bCfgOk := (fDwellMin_ms < fDwellMax_ms)
        AND NOT ((fQualityTarget <> fQualityTarget) OR ((fQualityTarget - fQualityTarget) <> (fQualityTarget - fQualityTarget)))
        AND (fQualityTarget >= DL_DW_TGT_LO) AND (fQualityTarget <= DL_DW_TGT_HI)
        AND (fDwellNominal_ms >= DL_DW_NOM_LO) AND (fDwellNominal_ms <= DL_DW_NOM_HI)
        AND (fTrimGain >= 0.0) AND (fTrimGain <= DL_DW_GAIN_HI)
        AND (fDwellRateMax_msS >= DL_DW_RATE_LO) AND (fDwellRateMax_msS <= DL_DW_RATE_HI);
IF NOT _bCfgOk THEN
    _bFaultLatch := TRUE;                           // 组态故障锁存 / Configuration fault latched
    eErr := DL_DW_CFG_BAD;                          // 故障级：组态非法 / Fault, bad configuration
    _eState := E_DL_DwellState.eFault;
END_IF

// 段 4｜质量可信闸（非有限即冻结微调，给定保持上次值）
_bQualityOk := NOT ((fSealQuality <> fSealQuality) OR ((fSealQuality - fSealQuality) <> (fSealQuality - fSealQuality)));
IF NOT _bQualityOk THEN
    eErr := DL_DW_QUAL_BAD;                         // 故障级：质量非有限，微调冻结 / Fault, the quality is not finite and the trim is frozen
    _eState := E_DL_DwellState.eFrozen;
END_IF

// 段 5｜微调积分（仅在运行、使能、组态与质量均可信时推进）
IF bEnable AND bRunning AND _bCfgOk AND _bQualityOk THEN
    _fErr := fQualityTarget - fSealQuality;         // 质量误差（正 = 质量偏低）/ Quality error, positive means poor sealing
    _fTrimWant := _fTrimWant + (_fErr * fTrimGain); // 期望微调分量积分 [ms] / Desired trim integrated
    // 先限速：单拍最大变化 = 变化率 × 代理任务周期
    _fTrimStep := fDwellRateMax_msS * DL_DW_TASK_S; // 本拍允许步长 [ms] / Allowed step of this scan
    _fTrimDelta := _fTrimWant - (_fDwellPrev - fDwellNominal_ms);   // 与上一拍的差 [ms] / Difference against the previous value
    IF _fTrimDelta > _fTrimStep THEN
        _fTrimDelta := _fTrimStep;                  // 正向限速 [ms] / Positive rate limit
    END_IF
    IF _fTrimDelta < (0.0 - _fTrimStep) THEN
        _fTrimDelta := 0.0 - _fTrimStep;            // 负向限速 [ms] / Negative rate limit
    END_IF
    _fDwellRaw := _fDwellPrev + _fTrimDelta;        // 限速后驻留 [ms] / Rate-limited dwell
    // 后钳制：把限速结果压进上下限，越限即触限并计数
    fDwellOut_ms := LIMIT(fDwellMin_ms, _fDwellRaw, fDwellMax_ms);
    IF ABS(fDwellOut_ms - _fDwellRaw) > 0.0001 THEN
        bAtLimit := TRUE;                           // 触限：给定被钳制 / At a bound, the setpoint was clamped
        eErr := DL_DW_LIMIT;                        // 信息级：触限钳制 / Info, clamped at a bound
        _eState := E_DL_DwellState.eAtLimit;
    ELSE
        _eState := E_DL_DwellState.eTrim;           // 正常微调 / Normal trimming
    END_IF
    _fTrimWant := fDwellOut_ms - fDwellNominal_ms;  // 反写分量（防积分饱和）[ms] / Anti-windup write-back
    IF ABS(_fTrimDelta) >= DL_DW_TRIM_EPS THEN
        uTrimCnt := uTrimCnt + 1;                   // 微调生效计数 +1 [次] / Effective trim count incremented
    END_IF
    _fDwellPrev := fDwellOut_ms;                    // 上一拍驻留快照 [ms] / Previous dwell snapshot
ELSE
    fDwellOut_ms := _fDwellPrev;                    // 冻结：保持上次给定 [ms] / Frozen, the previous setpoint is held
    IF _bQualityOk AND bEnable AND (NOT _bCfgOk) THEN
        eErr := DL_DW_CFG_BAD;                      // 故障级：组态非法保持 / Fault, the configuration error is held
    END_IF
END_IF

// 段 6｜微调分量出口与相位收口（ENUM + CASE + ELSE 兜底）
fDwellTrim_ms := _fTrimWant;                        // 微调分量出口 [ms] / Trim component output
CASE _eState OF
    E_DL_DwellState.eFrozen:
        bAtLimit := FALSE;                          // 冻结期不报触限 / No bound report while frozen
        IF bEnable AND bRunning AND _bCfgOk AND _bQualityOk THEN
            _eState := E_DL_DwellState.eTrim;       // 条件齐备：转微调 / Conditions met, go trimming
        END_IF
    E_DL_DwellState.eTrim:
        IF (NOT bRunning) OR (NOT bEnable) THEN
            _eState := E_DL_DwellState.eFrozen;     // 停机或失能：冻结 / Stopped or disabled, freeze
        END_IF
    E_DL_DwellState.eAtLimit:
        IF (NOT bRunning) OR (NOT bEnable) THEN
            _eState := E_DL_DwellState.eFrozen;
        END_IF
    E_DL_DwellState.eFault:
        eErr := DL_DW_CFG_BAD;                      // 故障级：组态非法保持 / Fault, the configuration error is held
        IF _bCfgOk AND (NOT bEnable) THEN
            _bFaultLatch := FALSE;                  // 组态修正且失能后解除 / Released after the configuration is fixed and the unit is disabled
            _eState := E_DL_DwellState.eFrozen;
        END_IF
    ELSE
        // 非法相位兜底（故障级）
        eErr := DL_DW_CFG_BAD;
        _bFaultLatch := TRUE;
        _eState := E_DL_DwellState.eFault;
END_CASE
IF eErr = 0 THEN
    eErr := DL_DW_READY;                            // 无事件回就绪码 / Ready code when nothing else applies
END_IF
END_FUNCTION_BLOCK

(* ---- FB_DL_SeasonMonthSched.st ---- *)
(*
  FB_DL_SeasonMonthSched  —  供暖/制冷季月度切换窗（月位图 + 切换滞回确认） / Season month schedule: heating/cooling bitmap with changeover hysteresis
  分类 Category : DL_Process
  版本 Version  : 1.0.0
  来源 Source   : t1-2-oscat-building — 楼宇季节切换族零检索深化
  溯源 Origin   : clean-room 实现，月位图语义公开借鉴 OSCAT 惯例，未复制任何源码行
  功能 Function : 1) 月度季节判据：uMonth（1..12）索引两幅 12 位月位图
                  （wHeatBmp 位 n-1 = 月 n 供暖 / wCoolBmp 位 n-1 = 月 n 制冷），
                  两位图均未命中 → 过渡季；
                  2) 切换滞回：目标季与当前季不一致 → eChgWait 相 tHyst 确认窗，
                  窗满提交切换，窗内目标季回撤即取消（eWait 相双出口，R98）；
                  3) 故障级三码独立：0382 位图交叠（同月双季，组态级锁存）/
                  0383 月值越界（uMonth > 12 判据不可信）/ 0384 ELSE 兜底；
                  4) 信息级三码：切供暖沿 / 切制冷沿 / 进过渡季沿；
                  5) 解除式全当拍量（R240 落地），逐 BOOL 标注见段 4。
  边界 Boundary : ① 位图判读前先做 uMonth 域闸（1..12），越界月不进移位判读
                  （移位量归一先于判据，R48 落地）；掩码用 SHL(WORD#1, 0..11)，
                  量域 0..11 < 16 结构性安全；
                  ② 位图交叠属静态组态错：锁存后季节出口保持当前季（冻结声明），
                  不随越界月漂移；
                  ③ 无 GVL 依赖：纯引脚输入输出，无外部变量引用，无物理 IO 地址。
  依赖 Depends  : Standard.library（TON / R_TRIG）
  码表 Error codes（Process 段 0005，窗口 0382~0384 / 04AA~04AC）:
    16#0005_0382 故障级：月位图交叠锁存（同月既供暖又制冷），锁存至 bReset
    16#0005_0383 故障级：月值越界锁存（uMonth > 12 判据不可信），锁存至 bReset
    16#0005_0384 故障级：相位落 ELSE 兜底或滞回窗域非法（tHyst <= 0，归并声明），锁存至 bReset
    16#0005_04AA 信息级：切换至供暖季沿
    16#0005_04AB 信息级：切换至制冷季沿
    16#0005_04AC 信息级：进入过渡季沿
  修订历史 Revision :
    2026-11-19  v1.0.0  R42 首版（批次 2 · 序号 2）
*)

TYPE E_DL_SmsSeason :
(
    eTrans  := 0,    // 过渡季：位图未命中 / Transition season
    eHeat   := 10,   // 供暖季 / Heating season
    eCool   := 20    // 制冷季 / Cooling season
);
END_TYPE

TYPE E_DL_SmsState :
(
    eIdle    := 0,   // 季节稳态：按当前季输出 / Steady season state
    eChgWait := 10,  // 切换确认：滞回窗计时 / Changeover confirm window
    eFault   := 90   // 故障：组态或月值锁定 / Fault, latched
);
END_TYPE

FUNCTION_BLOCK FB_DL_SeasonMonthSched
VAR_INPUT
    uMonth       : USINT := 1;        // 当前月 [1..12]，越界判 0383 / Current month
    wHeatBmp     : WORD := 16#0FC0;   // 供暖月位图，位 n-1 = 月 n 供暖 / Heating month bitmap
    wCoolBmp     : WORD := 16#003C;   // 制冷月位图，位 n-1 = 月 n 制冷 / Cooling month bitmap
    tHyst        : TIME := T#10M;     // 切换滞回确认窗 [ms]，域 > 0 / Changeover hysteresis window
    bReset       : BOOL := FALSE;     // 复位，上升沿清故障锁存 / Reset edge clears fault latch
END_VAR
VAR_OUTPUT
    eState       : E_DL_SmsState;     // 相位出口，段尾单点映射 / State outlet
    eSeason      : E_DL_SmsSeason;    // 当前季出口 / Current season outlet
    bHeatDemand  : BOOL;              // 供暖需求出口（供暖季电平）[-] / Heating demand outlet
    bCoolDemand  : BOOL;              // 制冷需求出口（制冷季电平）[-] / Cooling demand outlet
    bError       : BOOL;              // 故障锁存标志 / Fault latch flag
    nErrId       : UDINT;             // 事件码，0 = 无事件 / Event code
END_VAR
VAR
    tonHyst      : TON;               // 切换滞回确认窗（eChgWait 相独占），无条件刷新 / Hysteresis timer
    rtReset      : R_TRIG;            // 复位沿实例，无条件刷新 / Reset edge instance
    _eState      : E_DL_SmsState := E_DL_SmsState.eIdle;   // 内部相位，CASE 唯一写入目标 / Internal phase, the only CASE write target
    _eSeason     : E_DL_SmsSeason := E_DL_SmsSeason.eTrans;  // 内部季（CASE 唯一写入目标）/ Internal season
    _eTgtSeason  : E_DL_SmsSeason;    // 月位图判出目标季 / Bitmap-derived target season
    _wMask       : WORD;              // 当月掩码（SHL 结果）/ Current month mask
    _bHeatHit    : BOOL;              // 供暖位命中当拍量 [-] / Heating-bit hit flag
    _bCoolHit    : BOOL;              // 制冷位命中当拍量 [-] / Cooling-bit hit flag
    _bMonthBad   : BOOL;              // 月值越界当拍量 [-] / Month-out-of-range flag
    _bBmpOvl     : BOOL;              // 位图交叠当拍量（静态组态错逐月判出）[-] / Bitmap overlap flag
    _bFault      : BOOL;              // 故障锁存位（锁存量）/ Latched fault bit
    _uFault      : UDINT;             // 故障码锁存（锁存量）/ Latched fault code
    _uInfo       : UDINT;             // 信息码，每拍重算 / Transient info code
END_VAR

(* —— 段 0：定时器与沿实例无条件周期刷新（禁置于 IF/CASE 内） —— *)
_bMonthBad := (uMonth = 0) OR (uMonth > 12);             // 月值越界（当拍量）
IF NOT _bMonthBad THEN               // 域内才进移位判读（移位量 0..11 结构性安全）
    _wMask := SHL(WORD#1, UINT(uMonth) - UINT#1);        // 当月掩码（移位量归一后合法域）
    _bHeatHit := (wHeatBmp AND _wMask) <> WORD#0;        // 供暖位命中（当拍量）
    _bCoolHit := (wCoolBmp AND _wMask) <> WORD#0;        // 制冷位命中（当拍量）
    _bBmpOvl := _bHeatHit AND _bCoolHit;                 // 位图交叠（当拍量）
    IF _bHeatHit THEN
        _eTgtSeason := E_DL_SmsSeason.eHeat;             // 目标季：供暖
    ELSIF _bCoolHit THEN
        _eTgtSeason := E_DL_SmsSeason.eCool;             // 目标季：制冷
    ELSE
        _eTgtSeason := E_DL_SmsSeason.eTrans;            // 目标季：过渡
    END_IF
END_IF
rtReset(CLK := bReset);              // 复位沿（每拍必调）
tonHyst(IN := (_eState = E_DL_SmsState.eChgWait), PT := tHyst);  // 滞回窗（确认相独占）

(* —— 段 1：单拍量预清零（锁存量 _bFault/_uFault 不入清单，禁同拍抹除） —— *)
_uInfo := 16#0000_0000;             // 信息码每拍重算
nErrId := 16#0000_0000;             // 事件码缺省无事件

(* —— 段 2：复位沿 + 域闸锁存（判据当拍量） —— *)
IF rtReset.Q THEN                   // rtReset.Q = 当拍量
    _bFault := FALSE;               // 清故障锁存位
    _uFault := 16#0000_0000;        // 清故障锁存码
END_IF
IF _bBmpOvl THEN                    // 位图交叠（当拍量，静态组态错）
    _uFault := 16#0005_0382;        // 故障级：位图交叠锁存
    _bFault := TRUE;                // 故障标志与码位配对（R45）
END_IF
IF _bMonthBad THEN                  // 月值越界（当拍量）
    _uFault := 16#0005_0383;        // 故障级：月值越界锁存
    _bFault := TRUE;
END_IF
IF TIME_TO_DINT(tHyst) <= 0 THEN    // 滞回窗域闸（当拍量）
    _uFault := 16#0005_0384;        // 故障级：组态非法（归并 0384，码表声明）
    _bFault := TRUE;
END_IF

(* —— 段 3：故障解除式（R240 落地，逐 BOOL 标注）：
     rtReset.Q = 当拍量；NOT _bBmpOvl = 当拍量；NOT _bMonthBad = 当拍量。
     均不含锁存量（_bFault/_uFault），解除边真实可达（组态修正 + 月值恢复 + 复位沿）。 —— *)
IF rtReset.Q AND (NOT _bBmpOvl) AND (NOT _bMonthBad) THEN
    _bFault := FALSE;               // 清故障锁存位（锁存量，仅此当拍量解除沿可清）
    _uFault := 16#0000_0000;        // 清故障锁存码（锁存量，仅本当拍量解除沿可清）
    IF _eState = E_DL_SmsState.eFault THEN
        _eState := E_DL_SmsState.eIdle;     // 故障相迁出：回稳态
    END_IF
END_IF

(* —— 段 4：相位机（CASE 全覆盖 + ELSE 兜底） —— *)
CASE _eState OF

E_DL_SmsState.eIdle:
    IF (NOT _bFault) AND (_eTgtSeason <> _eSeason) THEN
        _eState := E_DL_SmsState.eChgWait;      // 目标季变更：进切换确认相
    END_IF

E_DL_SmsState.eChgWait:
    IF tonHyst.Q THEN                           // 出口 1：滞回窗满（事件量）
        CASE _eTgtSeason OF                     // 切换提交拍按目标季发信息沿（码表声明逐分支对齐）
            E_DL_SmsSeason.eHeat:
                _uInfo := 16#0005_04AA;         // 信息级：切换至供暖季沿
            E_DL_SmsSeason.eCool:
                _uInfo := 16#0005_04AB;         // 信息级：切换至制冷季沿
            E_DL_SmsSeason.eTrans:
                _uInfo := 16#0005_04AC;         // 信息级：进入过渡季沿
            ELSE
                _eState := E_DL_SmsState.eFault;    // 目标季非法兜底：进故障相（安全默认，不提交切换）/ Illegal target season fallback, enter fault, do not commit
                _bFault := TRUE;                    // 故障锁存与码位配对 / Fault latch paired with code
                _uFault := 16#0005_0384;            // 故障级：滞回窗域非法/兜底归并码 / Fault level, merged fallback code
        END_CASE
        IF NOT _bFault THEN                     // 兜底拍不提交切换（安全侧）/ Do not commit the switch in the fallback scan
            _eSeason := _eTgtSeason;                // 提交切换（锁存量级提交）
            _eState := E_DL_SmsState.eIdle;         // 回稳态相
        END_IF
    ELSIF _eTgtSeason = _eSeason THEN           // 出口 2：目标季回撤（前置条件消失，R98 双出口）
        _eState := E_DL_SmsState.eIdle;         // 取消切换：回稳态相
    END_IF

E_DL_SmsState.eFault:
    ;                                           // 故障相：季节出口冻结当前季（头注释②声明）
    (* 解除迁出在段 3 承载 *)

ELSE
    _uFault := 16#0005_0384;                // 故障级：非法相位兜底
    _bFault := TRUE;
    _eState := E_DL_SmsState.eFault;        // 强制回故障相

END_CASE

(* —— 段 6：出口单点映射（名实同源；锁存码回放，禁同拍抹除） —— *)
IF (_eSeason = E_DL_SmsSeason.eHeat) AND (NOT _bFault) THEN
    bHeatDemand := TRUE;            // 供暖需求（电平）
ELSE
    bHeatDemand := FALSE;           // 非供暖季强制 FALSE
END_IF
IF (_eSeason = E_DL_SmsSeason.eCool) AND (NOT _bFault) THEN
    bCoolDemand := TRUE;            // 制冷需求（电平）
ELSE
    bCoolDemand := FALSE;           // 非制冷季强制 FALSE
END_IF
IF _bFault THEN
    nErrId := _uFault;              // 故障锁存码回放
ELSE
    nErrId := _uInfo;               // 信息码
END_IF
bError := _bFault;                  // 故障标志与锁存位同源
eSeason := _eSeason;                // 季节出口单点映射
eState := _eState;                  // 相位出口单点映射

END_FUNCTION_BLOCK
